pHeader := iq_stEntry.pRxBuffer;
IF pHeader = 0 THEN
	RETURN;
END_IF
IF pHeader^.DeviceCount=0 OR pHeader^.DeviceCount>iq_stEntry.nMaxRecords THEN RETURN; END_IF
IF pHeader^.DeviceCount>(nPayloadBytes-SIZEOF(ST_MqttCommandHeader))/iq_stEntry.nElementSize THEN RETURN; END_IF
nRequiredBytes:=SIZEOF(ST_MqttCommandHeader)+pHeader^.DeviceCount*iq_stEntry.nElementSize;
IF nRequiredBytes>nPayloadBytes THEN RETURN; END_IF
nRecords := pHeader^.DeviceCount;		// 버퍼에 들어갈 수만큼 (위 검사로 실제 받은 레코드 수 이하)
q_nReceived := nRecords;		// [STD 21번 수정 2026-11-09: 받은 레코드 수]

(* 1부터 셈: 레코드가 0개면 돌지 않음 (0 - 1을 UDINT로 계산하면 넘쳐서 약 42억 번 돌게 됨) *)
FOR k := 1 TO nRecords DO
	pRecord := iq_stEntry.pRxBuffer;
	pRecord := pRecord + SIZEOF(ST_MqttCommandHeader) + (k - 1) * iq_stEntry.nElementSize;

	IF iq_stEntry.bIndexed THEN
		pIndex := pRecord + iq_stEntry.nIndexOffset;	// DeviceIndex 위치 (command는 SequenceNumber 뒤 4 B, config는 맨 앞) [2026-11-12]
		IF pIndex^ >= DEVICE_ID_BASE + iq_stEntry.nDeviceIdBase THEN
			nDev := pIndex^ - DEVICE_ID_BASE - iq_stEntry.nDeviceIdBase;
		ELSE
			nDev := iq_stEntry.nDeviceCapacity;	// 범위 밖 → 버림
		END_IF
	ELSE
		nDev := 0;							// 단일 레코드 (protection)
	END_IF

	IF nDev < iq_stEntry.nDeviceCapacity THEN
		pDest := iq_stEntry.pDestArray;
		pDest := pDest + nDev * iq_stEntry.nElementSize;
		MEMCPY(destAddr := pDest, srcAddr := pRecord, n := iq_stEntry.nElementSize);
		F_MqttDistribute := F_MqttDistribute + 1;
	END_IF
END_FOR

END_FUNCTION

// ---- 20_Module/Mqtt/FB_MqttPublish.TcPOU
FUNCTION_BLOCK FB_MqttPublish		// MQTT 발행 (브로커 1개): 장치 토픽·config echo 토픽을 1 s마다 발행, 로거 이벤트는 M_PublishLogger로 1건씩
VAR_INPUT
	i_nSiteId		: UDINT;
	i_sConnLabel	: STRING(10);	// 연결 구분 ('Cloud', 'local', 'Azure'). ClientId에만 씀
	i_sHost			: STRING(15);
	i_nPort			: UINT;
	i_sUserName		: STRING;
	i_sUserPassword	: STRING;	// 접속 값은 첫 호출 때 한 번 읽음
	i_sInstance		: STRING(4) := '';	// ClientId 뒤에 붙임. 이중화: 두 PLC가 같은 ClientId로 접속하면 브로커가 서로 끊으므로 PLC마다 다르게 ('-P', '-S')
	i_bPublish		: BOOL := TRUE;	// FALSE = 접속은 유지하고 발행만 안 함 (이중화: Active만 발행)
	i_astDeviceTable	: ARRAY[1..GVL_MQTT.DEVICE_TOPIC_COUNT] OF ST_MqttPubEntry;	// 장치 토픽 표 (FB_MqttMain.A_InitPublishTable)
	i_astConfigTable	: ARRAY[1..GVL_MQTT.CONFIG_TOPIC_COUNT] OF ST_MqttPubEntry;	// config echo 토픽 표
END_VAR
VAR
	_sSiteId			: STRING;
	_sClientId			: STRING;
	_sHost				: STRING(15);
	_nPort				: UINT;
	_sUserName			: STRING;
	_sUserPassword		: STRING;
	_asDeviceTopic		: ARRAY[1..GVL_MQTT.DEVICE_TOPIC_COUNT] OF STRING(80);
	_asConfigTopic		: ARRAY[1..GVL_MQTT.CONFIG_TOPIC_COUNT] OF STRING(80);
	_sLoggerTopic		: STRING(80);
	_fbClient			: FB_IotMqttClient;
	_fbQueue			: FB_IotMqttMessageQueue;
	_i					: UINT;
	_bSetParameter		: BOOL := TRUE;
	_bConnect			: BOOL := TRUE;
	_bPublished			: BOOL;
	_tonPeriod			: TON := (PT := T#1S);		// 발행 주기
END_VAR

IF _bSetParameter THEN
	_bSetParameter := FALSE;
	_sSiteId		:= UDINT_TO_STRING(i_nSiteId);
	_sHost			:= i_sHost;
	_nPort			:= i_nPort;
	_sClientId		:= CONCAT(CONCAT('dgspms/pub-', i_sConnLabel), CONCAT('/', _sSiteId));
	_sClientId		:= CONCAT(_sClientId, i_sInstance);
	_sUserName		:= i_sUserName;
	_sUserPassword	:= i_sUserPassword;
	(* 장치 토픽: dgspms/{solution}/{site_id}/{device_name} *)
	FOR _i := 1 TO GVL_MQTT.DEVICE_TOPIC_COUNT DO
		_asDeviceTopic[_i] := CONCAT(CONCAT(CONCAT('dgspms/', GVL_MQTT.SOLUTION_NAME), CONCAT('/', _sSiteId)),
									CONCAT('/', i_astDeviceTable[_i].sTopic));
	END_FOR
	(* config echo 토픽: dgspms/{solution}/{site_id}/config/{device_name} *)
	FOR _i := 1 TO GVL_MQTT.CONFIG_TOPIC_COUNT DO
		_asConfigTopic[_i] := CONCAT(CONCAT(CONCAT('dgspms/', GVL_MQTT.SOLUTION_NAME), CONCAT('/', _sSiteId)),
									CONCAT(CONCAT('/', i_astConfigTable[_i].sCategory), CONCAT('/', i_astConfigTable[_i].sTopic)));
	END_FOR

	(* 로거 토픽: dgspms/{solution}/{site_id}/{LOGGER_TOPIC} (주기 발행 아님. M_PublishLogger로 이벤트가 생길 때만) *)
	_sLoggerTopic := CONCAT(CONCAT(CONCAT('dgspms/', GVL_MQTT.SOLUTION_NAME), CONCAT('/', _sSiteId)), CONCAT('/', GVL_MQTT.LOGGER_TOPIC));

	_fbClient.sClientId		:= _sClientId;
	_fbClient.sUserName		:= _sUserName;
	_fbClient.sUserPassword	:= _sUserPassword;
	_fbClient.sHostName		:= _sHost;
	_fbClient.nHostPort		:= _nPort;
	_fbClient.sTopicPrefix	:= '';
	_fbClient.ipMessageQueue := _fbQueue;
END_IF

_fbClient.Execute(_bConnect);

IF _fbClient.bConnected AND i_bPublish THEN
	_tonPeriod(IN := TRUE);
	IF _tonPeriod.Q THEN
		_tonPeriod(IN := FALSE);
		FOR _i := 1 TO GVL_MQTT.DEVICE_TOPIC_COUNT DO
			IF i_astDeviceTable[_i].nDeviceCount > 0 THEN
			_bPublished := _fbClient.Publish(sTopic := _asDeviceTopic[_i],
						pPayload := i_astDeviceTable[_i].pStaging,
						nPayloadSize := i_astDeviceTable[_i].nStagingSize,
						eQos := TcIotMqttQos.AtMostOnceDelivery,
						bRetain := FALSE,
						bQueue := FALSE);
			END_IF
		END_FOR
		FOR _i := 1 TO GVL_MQTT.CONFIG_TOPIC_COUNT DO
			IF i_astConfigTable[_i].nDeviceCount > 0 THEN
			_bPublished := _fbClient.Publish(sTopic := _asConfigTopic[_i],
						pPayload := i_astConfigTable[_i].pStaging,
						nPayloadSize := i_astConfigTable[_i].nStagingSize,
						eQos := TcIotMqttQos.AtMostOnceDelivery,
						bRetain := FALSE,
						bQueue := FALSE);
			END_IF
		END_FOR
	END_IF
END_IF

METHOD M_PublishLogger : BOOL		// 로거 이벤트 1건 발행 (QoS 1, 반복 없음). 접속돼 있고 보냈으면 TRUE (FB_MqttMain.A_PublishLogger가 부름)
VAR_INPUT
	i_pPayload	: PVOID;		// ST_LoggerPublish_V1
	i_nSize		: UDINT;
END_VAR
M_PublishLogger := FALSE;
IF _bSetParameter OR NOT _fbClient.bConnected OR NOT i_bPublish THEN
	RETURN;		// 아직 접속 전: 큐에 남아 있다가 접속하면 나감. 발행 허가 없음(이중화 대기)도 보내지 않음
END_IF
M_PublishLogger := _fbClient.Publish(sTopic := _sLoggerTopic,
						pPayload := i_pPayload,
						nPayloadSize := i_nSize,
						eQos := TcIotMqttQos.AtLeastOnceDelivery,
						bRetain := FALSE,
						bQueue := FALSE);
END_METHOD

END_FUNCTION_BLOCK

// ---- 20_Module/Mqtt/Logger/FB_MqttLoggerListener.TcPOU
FUNCTION_BLOCK FB_MqttLoggerListener EXTENDS FB_ListenerBase2		// 로거 리스너: TwinCAT 이벤트 로거에 남은 PMS 이벤트를 받아 시각·문구를 큐에 쌓음 (로거 토픽 발행용. FB_MqttMain이 M_Cycle·M_GetPacket을 부름)
(* - FB_EventLog가 이벤트 로거에 남긴 것을 그대로 받는다 (메시지 1회, 알람 발생·해소). 기록하는 곳은 FB_EventLog 하나이고, 이 FB는 받아서 옮기기만 한다
   - 받는 이벤트 클래스: PmsSystem·PmsProt·PmsOutput·PmsSeq (TwinCAT 시스템 이벤트는 받지 않음). 구독은 클래스 단위(TC_EVENT_CLASSES)
   - 제어기 TwinCAT 런타임 3.1.4024.17 이상 필요 (FB_ListenerBase2). 낮으면 구독이 16#98110701(서비스 미지원)로 실패해 아무것도 받지 못함 (_hrSubscribe)
   - 문구: FB_RequestEventText로 비동기로 받는다 (UTF-8 → F_Utf8ToWstring). 해소는 앞에 '[해소] '.
     LOGGER_TEXT_MAX(100)자를 넘으면 99자 + '…'로 자르고 q_nTruncated를 센다 (문구 규칙: 인자를 채운 로그 문구 95자 이내, PMS_STD.md 7장)
   - 시각: 로거 기록 시각(UTC)을 현지 시각으로 바꾼다 (i_nUtcOffset, FB_MqttMain이 계산). 시간대를 아직 모르면 기다린다
   - 큐: LOGGER_QUEUE칸 링 버퍼. 브로커마다 M_GetPacket으로 다음 번호를 꺼내 간다. 밀려서 덮어쓰인 것은 건너뛰고 q_nLost
   - 본체는 부르지 않는다 (리스너 기반 FB). 매 스캔 M_Cycle을 부른다 *)
VAR_OUTPUT
	q_bSubscribed	: BOOL;		// 이벤트 로거 구독 중
	q_nReceived		: UDINT;	// 받은 이벤트 수 (= 마지막 이벤트 번호)
	q_nTruncated	: UDINT;	// LOGGER_TEXT_MAX를 넘어 자른 수 (문구 규칙 위반: 문구 틀·인자를 줄일 것)
	q_nTextError	: UDINT;	// 문구를 못 받아 대체 문구를 쓴 수
	q_nLost			: UDINT;	// 브로커가 밀려 보내지 못하고 덮어쓰인 수 (브로커 합)
END_VAR
VAR CONSTANT
	TEXT_TIMEOUT	: ULINT := 50000000;	// 문구 요청 제한 5 s (100 ns 단위). 넘으면 대체 문구
	SUBSCRIBE_RETRY	: UINT := 100;			// 구독 실패 뒤 다시 시도까지 M_Cycle 호출 수 (MqttTask 10 ms × 100 = 1 s)
	CLEARED_MARK	: WSTRING(7) := "[해소] ";	// 알람 해소 표시 (5자)
END_VAR
VAR
	_fbFilter		: FB_TcEventFilter;
	_hrSubscribe	: HRESULT;
	_hrExecute		: HRESULT;
	_nSubscribeWait	: UINT;
	_nUtcOffset		: LINT;		// 현지 시각 − UTC (100 ns). M_Cycle 입력
	_bTimeValid		: BOOL;
	_nWriteNo		: UDINT;	// 마지막으로 넣은 이벤트 번호
	_astSlot		: ARRAY[1..GVL_MQTT.LOGGER_QUEUE] OF ST_LoggerSlot;
	_afbText		: ARRAY[1..GVL_MQTT.LOGGER_QUEUE] OF FB_RequestEventText;	// 칸마다 하나 (한 스캔에 여러 이벤트가 와도 요청이 겹치지 않게)
	{attribute 'TcEncoding' := 'UTF-8'}
	_sText			: STRING(511);		// 받은 문구 (UTF-8. 한글 95자 ≈ 285 byte)
	_wsText			: WSTRING(255);
	_k				: UINT;
	_nNow			: ULINT;
END_VAR

(* 본체는 쓰지 않는다. M_Cycle을 부른다 *)

METHOD M_Cycle		// 매 스캔 (MqttTask): 구독 → 이벤트 받기(콜백이 큐에 넣음) → 칸마다 문구·시각 채우기
VAR_INPUT
	i_nUtcOffset	: LINT;		// 현지 시각 − UTC (100 ns 단위)
	i_bTimeValid	: BOOL;		// i_nUtcOffset을 믿을 수 있음 (현지 시각을 얻음)
END_VAR
_nUtcOffset	:= i_nUtcOffset;
_bTimeValid	:= i_bTimeValid;

(* 1. 구독 (처음, 실패하면 SUBSCRIBE_RETRY 호출 뒤 다시) *)
IF NOT THIS^.bSubscribed THEN
	IF _nSubscribeWait = 0 THEN
		(* 클래스 단위 (TC_EVENT_CLASSES): 클래스 안의 이벤트를 추가·삭제·이름 변경해도 고치지 않음. 새 이벤트 클래스를 만들면 여기에 한 줄 *)
		_fbFilter.Clear().EventClass.EqualTo(TC_EVENT_CLASSES.PmsSystem)
			.OR_OP().EventClass.EqualTo(TC_EVENT_CLASSES.PmsProt)
			.OR_OP().EventClass.EqualTo(TC_EVENT_CLASSES.PmsOutput)
			.OR_OP().EventClass.EqualTo(TC_EVENT_CLASSES.PmsSeq);
		_hrSubscribe := THIS^.Subscribe2(_fbFilter);
		_nSubscribeWait := SUBSCRIBE_RETRY;
	ELSE
		_nSubscribeWait := _nSubscribeWait - 1;
	END_IF
END_IF
q_bSubscribed := THIS^.bSubscribed;

(* 2. 이벤트 받기: 이 안에서 OnMessageSent·OnAlarmRaised·OnAlarmCleared가 불려 큐에 넣고 문구를 요청함 *)
_hrExecute := THIS^.Execute();

(* 3. 칸마다: 문구가 오면 받고, 시간대를 알면 시각 문자열을 만들어 발행 준비 *)
_nNow := F_GetSystemTime();
FOR _k := 1 TO GVL_MQTT.LOGGER_QUEUE DO
	IF _astSlot[_k].bRequesting THEN
		IF _afbText[_k].bError OR (_nNow - _astSlot[_k].nRequestStart) > TEXT_TIMEOUT THEN
			q_nTextError := q_nTextError + 1;
			M_SetText(i_nSlot := _k, i_wsText := WCONCAT("로그 문구를 가져오지 못함: 이벤트 ID ", TO_WSTRING(_astSlot[_k].nEventId)));
		ELSIF NOT _afbText[_k].bBusy THEN
			_sText := '';
			_afbText[_k].GetString(_sText, SIZEOF(_sText));
			M_SetText(i_nSlot := _k, i_wsText := F_Utf8ToWstring(i_pSrc := ADR(_sText), i_nSrcSize := SIZEOF(_sText)));
		END_IF
	END_IF
	IF _astSlot[_k].bTextDone AND NOT _astSlot[_k].bReady AND _bTimeValid THEN
		_astSlot[_k].sTime	:= M_TimeText(_astSlot[_k].nTimestamp);
		_astSlot[_k].bReady	:= TRUE;
	END_IF
END_FOR
END_METHOD

METHOD M_GetPacket : BOOL		// 브로커 하나가 보낼 다음 이벤트 패킷. TRUE면 iq_stPacket을 채움 (보낸 뒤 부르는 쪽이 iq_nNext를 1 올림)
VAR_INPUT
	i_nSiteId	: UDINT;
END_VAR
VAR_IN_OUT
	iq_nNext	: UDINT;				// 이 브로커가 다음에 보낼 이벤트 번호 (1부터)
	iq_stPacket	: ST_LoggerPublish_V1;
END_VAR
VAR
	k			: UINT;
	nOldest		: UDINT;
	nBytes		: UDINT;
END_VAR
M_GetPacket := FALSE;
IF iq_nNext = 0 THEN
	iq_nNext := 1;
END_IF
IF _nWriteNo < iq_nNext THEN
	RETURN;		// 새 이벤트 없음
END_IF

(* 큐 칸 수보다 많이 밀렸으면 덮어쓰인 것은 건너뜀 *)
IF _nWriteNo - iq_nNext >= UINT_TO_UDINT(GVL_MQTT.LOGGER_QUEUE) THEN
	nOldest		:= _nWriteNo - UINT_TO_UDINT(GVL_MQTT.LOGGER_QUEUE) + 1;
	q_nLost		:= q_nLost + (nOldest - iq_nNext);
	iq_nNext	:= nOldest;
END_IF

k := M_SlotOf(iq_nNext);
IF _astSlot[k].nNo <> iq_nNext OR NOT _astSlot[k].bReady THEN
	RETURN;		// 문구·시각을 아직 받는 중
END_IF

(* 매번 비우고 채움: 짧은 문구의 null 뒤에 지난 문구가 남지 않게.
   문자열은 대입(:=)하지 않고 길이 + null만 MEMCPY: 문자열 대입은 선언 크기 전체를 복사해서,
   큐 칸을 돌려 쓰는 동안 null 뒤에 남은 옛 문구까지 패킷에 들어감 (PC 도구 재pack 비교에서 "불일치"로 보임) *)
MEMSET(destAddr := ADR(iq_stPacket), fillByte := 0, n := SIZEOF(iq_stPacket));
iq_stPacket.Header.HeaderVersion	:= GVL_MQTT.HEADER_VERSION;
iq_stPacket.Header.DeviceVersion	:= GVL_MQTT.LOGGER_VERSION;
iq_stPacket.Header.SiteId			:= i_nSiteId;
nBytes := INT_TO_UDINT(LEN(_astSlot[k].sTime)) + 1;
IF nBytes > SIZEOF(iq_stPacket.Header.TimeStamp) THEN
	nBytes := SIZEOF(iq_stPacket.Header.TimeStamp);
END_IF
MEMCPY(destAddr := ADR(iq_stPacket.Header.TimeStamp), srcAddr := ADR(_astSlot[k].sTime), n := nBytes);
nBytes := (INT_TO_UDINT(WLEN(_astSlot[k].wsText)) + 1) * 2;
IF nBytes > SIZEOF(iq_stPacket.Contents) THEN
	nBytes := SIZEOF(iq_stPacket.Contents);
END_IF
MEMCPY(destAddr := ADR(iq_stPacket.Contents), srcAddr := ADR(_astSlot[k].wsText), n := nBytes);
M_GetPacket := TRUE;
END_METHOD

METHOD OnMessageSent : HRESULT		// 메시지 1건 (FB_LogMsg) → 큐
VAR_INPUT
	fbEvent	: REFERENCE TO FB_TcEvent;
END_VAR
M_Push(i_fbEvent := fbEvent, i_bCleared := FALSE);
OnMessageSent := S_OK;		// S_OK여야 이번 스캔에 다음 콜백을 계속 받음
END_METHOD

METHOD OnAlarmRaised : HRESULT		// 알람 발생 (FB_LogAlarm) → 큐
VAR_INPUT
	fbEvent	: REFERENCE TO FB_TcEvent;
END_VAR
M_Push(i_fbEvent := fbEvent, i_bCleared := FALSE);
OnAlarmRaised := S_OK;		// S_OK여야 이번 스캔에 다음 콜백을 계속 받음
END_METHOD

METHOD OnAlarmCleared : HRESULT		// 알람 해소 → 큐 ('[해소] ' 표시)
VAR_INPUT
	fbEvent	: REFERENCE TO FB_TcEvent;
END_VAR
M_Push(i_fbEvent := fbEvent, i_bCleared := TRUE);
OnAlarmCleared := S_OK;		// S_OK여야 이번 스캔에 다음 콜백을 계속 받음
END_METHOD

METHOD OnAlarmConfirmed : HRESULT		// 쓰지 않음
VAR_INPUT
	fbEvent	: REFERENCE TO FB_TcEvent;
END_VAR
OnAlarmConfirmed := S_OK;		// 확인(Confirm)은 쓰지 않음 (알람을 확인 없이 만듦)
END_METHOD

METHOD PRIVATE M_Push		// 받은 이벤트를 큐 다음 칸에 넣고 문구를 요청 (콜백이 부름). 큐가 차면 가장 오래된 칸을 덮어씀
VAR_INPUT
	i_fbEvent	: REFERENCE TO FB_TcEvent;
	i_bCleared	: BOOL;
END_VAR
VAR
	k			: UINT;
END_VAR
_nWriteNo	:= _nWriteNo + 1;
q_nReceived	:= _nWriteNo;
k := M_SlotOf(_nWriteNo);

_astSlot[k].nNo				:= _nWriteNo;
_astSlot[k].nTimestamp		:= i_fbEvent.nTimestamp;
_astSlot[k].nEventId		:= i_fbEvent.nEventId;
_astSlot[k].bCleared		:= i_bCleared;
_astSlot[k].bRequesting		:= TRUE;
_astSlot[k].nRequestStart	:= F_GetSystemTime();
_astSlot[k].bTextDone		:= FALSE;
_astSlot[k].bReady			:= FALSE;
_astSlot[k].sTime			:= '';
_astSlot[k].wsText			:= "";

(* 문구는 비동기로 옴 (M_Cycle에서 받음). 인자는 요청할 때 넘김 (콜백 밖에서는 i_fbEvent를 쓸 수 없음) *)
_afbText[k].Request(eventClass := i_fbEvent.EventClass, nEventId := i_fbEvent.nEventId,
					nLangId := GVL_MQTT.LOGGER_LANG_ID, ipArgs := i_fbEvent.ipArguments);
END_METHOD

METHOD PRIVATE M_SetText		// 받은 문구를 칸에 넣음: 해소 표시를 붙이고 LOGGER_TEXT_MAX자로 맞춤
VAR_INPUT
	i_nSlot		: UINT;
	i_wsText	: WSTRING(255);
END_VAR
_wsText := i_wsText;
IF _astSlot[i_nSlot].bCleared THEN
	_wsText := WCONCAT(CLEARED_MARK, _wsText);
END_IF
IF WLEN(_wsText) > GVL_MQTT.LOGGER_TEXT_MAX THEN
	_wsText := WCONCAT(WLEFT(_wsText, GVL_MQTT.LOGGER_TEXT_MAX - 1), "…");
	q_nTruncated := q_nTruncated + 1;
END_IF
_astSlot[i_nSlot].wsText		:= _wsText;
_astSlot[i_nSlot].bRequesting	:= FALSE;
_astSlot[i_nSlot].bTextDone		:= TRUE;
END_METHOD

METHOD PRIVATE M_SlotOf : UINT		// 이벤트 번호 → 큐 칸 (1..LOGGER_QUEUE)
VAR_INPUT
	i_nNo	: UDINT;
END_VAR
M_SlotOf := UDINT_TO_UINT(((i_nNo - 1) MOD UINT_TO_UDINT(GVL_MQTT.LOGGER_QUEUE)) + 1);
END_METHOD

METHOD PRIVATE M_TimeText : STRING(23)		// 로거 시각(FILETIME, UTC) → 현지 시각 문자열
VAR_INPUT
	i_nFileTime	: ULINT;
END_VAR
VAR
	nLocal		: ULINT;
	stFileTime	: T_FILETIME;
END_VAR
nLocal := LINT_TO_ULINT(ULINT_TO_LINT(i_nFileTime) + _nUtcOffset);
MEMCPY(destAddr := ADR(stFileTime), srcAddr := ADR(nLocal), n := SIZEOF(stFileTime));
M_TimeText := F_MqttTimeText(FILETIME_TO_SYSTEMTIME(stFileTime));
END_METHOD

END_FUNCTION_BLOCK

// ---- 20_Module/Mqtt/Logger/F_Utf8ToWstring.TcPOU
FUNCTION F_Utf8ToWstring : WSTRING(255)		// UTF-8 바이트(0에서 끝남) → WSTRING(UTF-16). 255자에서 자름. 4바이트 문자(이모지 등)·잘못된 바이트는 U+FFFD 한 글자
(* 이벤트 로거 문구(FB_RequestEventText.GetString)는 UTF-8 STRING으로만 받을 수 있어서 쓴다.
   한글(U+AC00~)은 UTF-8 3바이트 → UTF-16 한 칸 *)
VAR_INPUT
	i_pSrc		: PVOID;				// UTF-8 문자열 시작 주소 (STRING 변수의 ADR)
	i_nSrcSize	: UDINT;				// 그 버퍼 크기 (byte, SIZEOF). 0을 만나면 그 앞에서 끝
END_VAR
VAR CONSTANT
	MAX_SRC		: UDINT := 1024;		// 읽는 최대 바이트
	MAX_CHARS	: UINT := 255;
	BAD_CHAR	: WORD := 16#FFFD;
END_VAR
VAR
	pSrc		: POINTER TO ARRAY[0..1023] OF BYTE;	// MAX_SRC
	wsOut		: WSTRING(255);
	pOut		: POINTER TO ARRAY[0..255] OF WORD;		// wsOut (MAX_CHARS + null)
	nSize		: UDINT;
	i			: UDINT;
	nChars		: UINT;
	nLen		: UDINT;
	b0			: BYTE;
	b1			: BYTE;
	b2			: BYTE;
	wChar		: WORD;
END_VAR

F_Utf8ToWstring := "";
IF i_pSrc = 0 THEN
	RETURN;
END_IF
pSrc	:= i_pSrc;
pOut	:= ADR(wsOut);
nSize	:= MIN(i_nSrcSize, MAX_SRC);
i		:= 0;
nChars	:= 0;

WHILE i < nSize AND nChars < MAX_CHARS DO
	b0 := pSrc^[i];
	IF b0 = 0 THEN
		EXIT;
	END_IF
	wChar	:= BAD_CHAR;
	nLen	:= 1;
	IF b0 < 16#80 THEN							// 1바이트 (ASCII)
		wChar := BYTE_TO_WORD(b0);
	ELSIF (b0 AND 16#E0) = 16#C0 THEN			// 2바이트
		IF i + 1 < nSize THEN
			b1 := pSrc^[i + 1];
			IF (b1 AND 16#C0) = 16#80 THEN
				wChar	:= SHL(BYTE_TO_WORD(b0 AND 16#1F), 6) OR BYTE_TO_WORD(b1 AND 16#3F);
				nLen	:= 2;
			END_IF
		END_IF
	ELSIF (b0 AND 16#F0) = 16#E0 THEN			// 3바이트 (한글 등)
		IF i + 2 < nSize THEN
			b1 := pSrc^[i + 1];
			b2 := pSrc^[i + 2];
			IF (b1 AND 16#C0) = 16#80 AND (b2 AND 16#C0) = 16#80 THEN
				wChar	:= SHL(BYTE_TO_WORD(b0 AND 16#0F), 12) OR SHL(BYTE_TO_WORD(b1 AND 16#3F), 6) OR BYTE_TO_WORD(b2 AND 16#3F);
				nLen	:= 3;
			END_IF
		END_IF
	ELSIF (b0 AND 16#F8) = 16#F0 THEN			// 4바이트 → U+FFFD 한 글자
		nLen := 4;
	END_IF
	pOut^[nChars]	:= wChar;
	nChars			:= nChars + 1;
	i				:= i + nLen;
END_WHILE
pOut^[nChars] := 0;
F_Utf8ToWstring := wsOut;

END_FUNCTION

// ---- 20_Module/Mqtt/F_MqttTimeText.TcPOU
FUNCTION F_MqttTimeText : STRING(23)		// 시각 → 'YYYY-MM-DD hh:mm:ss.xxx' (MQTT 헤더 TimeStamp 형식, 23자). FB_MqttMain(발행 헤더)·FB_MqttLoggerListener(로거 시각)가 같이 씀
VAR_INPUT
	i_stTime	: TIMESTRUCT;
END_VAR

(* Tc2_Utilities SYSTEMTIME_TO_STRING 형식은 'YYYY-MM-DD-hh:mm:ss.xxx' → 11번째 글자 '-'를 공백으로 *)
F_MqttTimeText := REPLACE(SYSTEMTIME_TO_STRING(i_stTime), ' ', 1, 11);

END_FUNCTION

// ---- 20_Module/Mqtt/FB_EmsCommand.TcPOU
FUNCTION_BLOCK FB_EmsCommand		// 명령 핸들러 (MqttTask): 받은 EMS command 레코드 → Std 명령 (PCS·BMS 상태 명령, 충전·방전 P 지령)
(* - 받은 레코드의 CommandType이 0이 아니면 한 번 해석하고 0으로 지운다 (같은 레코드를 다시 실행하지 않음)
   - 새 명령마다 번호(nSeq, anPcsPSeq)를 1 올린다. 받는 쪽(FB_SrcEms)은 번호 변화로 새 명령을 안다
   - 결과 q_stCmd는 지금까지 받은 명령 전체(마지막 값 유지). 바뀐 스캔에만 q_bChanged가 켜지고, PRG_Mqtt가 GVL_IF에 올린다
   - 받은 레코드 배열은 0부터 (GVL_MQTT 수신 배열 칸 = 레코드 DeviceIndex − 1, F_MqttDistribute.DEVICE_ID_BASE = 1). 결과는 Std 규칙대로 1부터 (칸 = DeviceIndex)
   - 이상한 값(NaN·무한대·절댓값이 MAX_VALUE 초과)의 P 지령은 버리고 센다. NaN은 비교하면 PLC가 멈추므로 F_IsFinite(비트)로 먼저 거른다. 정격 대비 상한은 코어 명령 필터(g_stCmdFilter)가 다시 거른다
   PCS CommandType: 1 Run, 2 Stop, 3 Standby, 4 충전(Value kW), 5 방전(Value kW), 6 비상정지, 7 리셋
   BAT CommandType: 1 접촉기 투입(Close), 2 개방(Open), 3 비상정지, 4 리셋, 11 랙 컨택터 닫기, 12 랙 컨택터 열기 (Value = 랙 번호 1~)
   5 시스템(랙 전체 40013) 연결, 6 차단, 7 충전 컨택터(40014) 닫기, 8 열기, 9 방전 컨택터(40015) 닫기, 10 열기 → astBatCtl [2026-11-13]
   (인터페이스 100.Command) *)
VAR_INPUT
	i_nRxCount			: UDINT;	// command 메시지 수신 누계 (브로커 3개 합)
END_VAR
VAR_IN_OUT
	iq_astPcsCommand	: ARRAY[0..GVL_PARAM.PCS_COUNT-1] OF ST_MqttCommand_Rx;	// GVL_MQTT.g_astPcsCommand
	iq_astBatCommand	: ARRAY[0..GVL_PARAM.BMS_COUNT-1] OF ST_MqttCommand_Rx;	// GVL_MQTT.g_astBatCommand
END_VAR
VAR_OUTPUT
	q_stCmd				: ST_IfEmsCmd;	// 지금까지 받은 명령
	q_bChanged			: BOOL;			// 이번 스캔에 q_stCmd가 바뀜
	q_nUnknownCount		: UDINT;		// 모르는 CommandType을 받은 횟수
	q_nBadValueCount	: UDINT;		// 이상한 값의 P 지령을 버린 횟수
END_VAR
VAR CONSTANT
	MAX_VALUE			: REAL := 1.0E7;	// kW. 이보다 크면 이상값
END_VAR
VAR
	_i					: UINT;
	_n					: UINT;
	_ePcsCmd			: E_PcsCmd;
	_eBatCmd			: E_BatCmd;
	_bP					: BOOL;
	_fP					: REAL;
	_bValueOk			: BOOL;		// 받은 Value가 보통 숫자 (NaN·무한대 아님)
END_VAR

q_bChanged := FALSE;

// 명령이 없는 메시지도 '살아 있음'으로 셈
IF i_nRxCount <> q_stCmd.nRxCount THEN
	q_stCmd.nRxCount := i_nRxCount;
	q_bChanged := TRUE;
END_IF

(* PCS *)
FOR _i := 0 TO GVL_PARAM.PCS_COUNT - 1 DO
	IF iq_astPcsCommand[_i].CommandType <> 0 THEN
		_n := _i + 1;
		_ePcsCmd	:= E_PcsCmd.None;
		_bP			:= FALSE;
		_bValueOk	:= F_IsFinite(iq_astPcsCommand[_i].Value);	// NaN은 크기 비교·ABS 전에 비트로 거름 (비교하면 PLC가 멈춤)
		CASE iq_astPcsCommand[_i].CommandType OF
			1:	_ePcsCmd := E_PcsCmd.Run;
			2:	_ePcsCmd := E_PcsCmd.Stop;
			3:	_ePcsCmd := E_PcsCmd.Standby;
			4:	_bP := TRUE;	IF _bValueOk THEN _fP := -ABS(iq_astPcsCommand[_i].Value); END_IF	// 충전
			5:	_bP := TRUE;	IF _bValueOk THEN _fP := ABS(iq_astPcsCommand[_i].Value); END_IF		// 방전
			6:	_ePcsCmd := E_PcsCmd.EStop;
			7:	_ePcsCmd := E_PcsCmd.Reset;
		ELSE
			q_nUnknownCount := q_nUnknownCount + 1;
		END_CASE
		// P 지령 값 거르기: 보통 숫자가 아니거나 너무 크면 버림 (크기 비교는 보통 숫자일 때만)
		IF _bP THEN
			IF NOT _bValueOk THEN
				_bP := FALSE;
				q_nBadValueCount := q_nBadValueCount + 1;
			ELSIF ABS(iq_astPcsCommand[_i].Value) > MAX_VALUE THEN
				_bP := FALSE;
				q_nBadValueCount := q_nBadValueCount + 1;
			END_IF
		END_IF
		IF _ePcsCmd <> E_PcsCmd.None THEN
			q_stCmd.astPcs[_n].eCmd := _ePcsCmd;
			q_stCmd.astPcs[_n].nSeq := q_stCmd.astPcs[_n].nSeq + 1;
			q_bChanged := TRUE;
		END_IF
		IF _bP THEN
			q_stCmd.afPcsP[_n]		:= _fP;
			q_stCmd.anPcsPSeq[_n]	:= q_stCmd.anPcsPSeq[_n] + 1;
			q_bChanged := TRUE;
		END_IF
		iq_astPcsCommand[_i].CommandType := 0;		// 처리 완료
	END_IF
END_FOR

(* BAT (BMS) *)
FOR _i := 0 TO GVL_PARAM.BMS_COUNT - 1 DO
	IF iq_astBatCommand[_i].CommandType <> 0 THEN
		_n := _i + 1;
		_eBatCmd := E_BatCmd.None;
		CASE iq_astBatCommand[_i].CommandType OF
			1:	_eBatCmd := E_BatCmd.Close;
			2:	_eBatCmd := E_BatCmd.Open;
			3:	_eBatCmd := E_BatCmd.EStop;
			4:	_eBatCmd := E_BatCmd.Reset;
			5..10:	// 컨택터 하나씩 (FB_BmsContactorCommand가 번호를 해석) [2026-11-13]
				q_stCmd.astBatCtl[_n].nSeq := q_stCmd.astBatCtl[_n].nSeq + 1;
				q_stCmd.astBatCtl[_n].nType := UDINT_TO_UINT(iq_astBatCommand[_i].CommandType);
				q_bChanged := TRUE;
			11, 12:	// 랙 컨택터 닫기·열기. Value = 랙 번호 (정수가 아니거나 범위 밖이면 0 → FB_BmsRackCommand가 거절)
				q_stCmd.astBatRack[_n].nSeq := q_stCmd.astBatRack[_n].nSeq + 1;
				q_stCmd.astBatRack[_n].bClose := iq_astBatCommand[_i].CommandType = 11;
				IF iq_astBatCommand[_i].Value >= 1.0 AND iq_astBatCommand[_i].Value <= 16.0
					AND iq_astBatCommand[_i].Value = UINT_TO_REAL(REAL_TO_UINT(iq_astBatCommand[_i].Value)) THEN
					q_stCmd.astBatRack[_n].nRack := REAL_TO_UINT(iq_astBatCommand[_i].Value);
				ELSE
					q_stCmd.astBatRack[_n].nRack := 0;
				END_IF
				q_bChanged := TRUE;
		ELSE
			q_nUnknownCount := q_nUnknownCount + 1;
		END_CASE
		IF _eBatCmd <> E_BatCmd.None THEN
			q_stCmd.astBat[_n].eCmd := _eBatCmd;
			q_stCmd.astBat[_n].nSeq := q_stCmd.astBat[_n].nSeq + 1;
			q_bChanged := TRUE;
		END_IF
		iq_astBatCommand[_i].CommandType := 0;		// 처리 완료
	END_IF
END_FOR

END_FUNCTION_BLOCK

// ---- 10_Core/02_Util/F_IsFinite.TcPOU
FUNCTION F_IsFinite : BOOL		// 실수가 보통 숫자인가 (NaN·무한대가 아님). 비트로만 봄
// NaN을 크기 비교(<, >, <=, >=)하면 부동소수점 예외(SSE invalid operation)로 PLC가 멈춤 → 바깥에서 온 실수는 비교하기 전에 이것으로 먼저 거름
VAR_INPUT
	i_fValue	: REAL;
END_VAR
VAR
	pBits		: POINTER TO DWORD;
END_VAR

pBits := ADR(i_fValue);
F_IsFinite := (pBits^ AND 16#7F800000) <> 16#7F800000;		// 지수 비트가 모두 1이면 NaN 또는 무한대

END_FUNCTION

// ---- 20_Module/Mqtt/FB_EmsCmdGate.TcPOU
FUNCTION_BLOCK FB_EmsCmdGate		// EMS command 레코드 앞단: 같은 SequenceNumber 버리기 + Delay(ms)만큼 기다렸다가 내보내기
(* EMS command 레코드 중복 방지·지연 실행 (⑤출력 앞단 / 장치: PCS·BAT·UPS 명령 공통). 2026-11-12.
   기반 없음(신규).
   변경: 없음
   부호·단위: Delay ms. 명세: C:\gil\UPS\명세서\UPS_명세서.md WR-CMD-01, 인터페이스 100.Command (SequenceNumber·Delay)
   - 수신 배열(GVL_MQTT.g_ast*Command, 칸 = DeviceIndex-1)을 그대로 받아, 명령 핸들러(FB_EmsCommand, PRG_Mqtt UPS 칸)보다 먼저 부른다
   - 새 레코드(CommandType<>0)의 SequenceNumber가 그 칸에서 마지막으로 받은 번호와 같으면 버린다 (0은 거르지 않음)
   - Delay = 0이면 그대로 두어 이번 스캔에 처리된다. Delay > 0이면 레코드를 빼서 보관하고, 시간이 되면 그 칸에 다시 넣는다
   - 보관 중에 같은 칸에 새 명령이 오면 보관한 명령은 버리고 새 명령을 따른다 (마지막 명령이 우선)
   - Delay가 MAX_DELAY_MS를 넘으면 버린다
   - 재시작하면 마지막 번호와 보관 명령은 없어진다 (보관 중이던 명령은 실행하지 않음) *)
VAR_IN_OUT
	iq_astRec			: ARRAY[*] OF ST_MqttCommand_Rx;	// 수신 배열 (0부터, 칸 = DeviceIndex-1)
END_VAR
VAR_OUTPUT
	q_nDupCount			: UDINT;	// 같은 SequenceNumber라 버린 수
	q_nDelayedCount		: UDINT;	// Delay 때문에 보관한 수
	q_nReplacedCount	: UDINT;	// 보관 중 새 명령이 와서 버린 보관 명령 수
	q_nBadDelayCount	: UDINT;	// Delay가 너무 커서 버린 수
	q_nPendingCount		: UDINT;	// 지금 보관 중인 명령 수
END_VAR
VAR CONSTANT
	MAX_SLOTS			: DINT := 16;			// 다룰 수 있는 칸 수 (PCS·BMS·UPS 대수보다 커야 함)
	MAX_DELAY_MS		: UDINT := 3600000;		// 1시간
END_VAR
VAR
	_anLastSeq			: ARRAY[0..15] OF UDINT;
	_astPend			: ARRAY[0..15] OF ST_MqttCommand_Rx;
	_abPend				: ARRAY[0..15] OF BOOL;
	_atStart			: ARRAY[0..15] OF TIME;
	_tNow				: TIME;
	_i					: DINT;
	_s					: DINT;
END_VAR

_tNow := TIME();
q_nPendingCount := 0;
FOR _i := LOWER_BOUND(iq_astRec, 1) TO UPPER_BOUND(iq_astRec, 1) DO
	_s := _i - LOWER_BOUND(iq_astRec, 1);
	IF _s >= MAX_SLOTS THEN
		EXIT;
	END_IF
	IF iq_astRec[_i].CommandType <> 0 THEN
		IF iq_astRec[_i].SequenceNumber <> 0 AND iq_astRec[_i].SequenceNumber = _anLastSeq[_s] THEN
			iq_astRec[_i].CommandType := 0;		// 같은 명령이 다시 옴
			q_nDupCount := q_nDupCount + 1;
		ELSE
			_anLastSeq[_s] := iq_astRec[_i].SequenceNumber;
			IF _abPend[_s] THEN
				_abPend[_s] := FALSE;			// 새 명령이 기다리던 명령을 대신함
				q_nReplacedCount := q_nReplacedCount + 1;
			END_IF
			IF iq_astRec[_i].Delay > MAX_DELAY_MS THEN
				iq_astRec[_i].CommandType := 0;
				q_nBadDelayCount := q_nBadDelayCount + 1;
			ELSIF iq_astRec[_i].Delay > 0 THEN
				_astPend[_s] := iq_astRec[_i];
				_abPend[_s] := TRUE;
				_atStart[_s] := _tNow;
				iq_astRec[_i].CommandType := 0;	// 시간이 될 때까지 핸들러가 못 보게 함
				q_nDelayedCount := q_nDelayedCount + 1;
			END_IF
		END_IF
	ELSIF _abPend[_s] AND (_tNow - _atStart[_s]) >= UDINT_TO_TIME(_astPend[_s].Delay) THEN
		iq_astRec[_i] := _astPend[_s];			// 시간이 됨: 이번 스캔에 핸들러가 처리
		iq_astRec[_i].Delay := 0;
		_abPend[_s] := FALSE;
	END_IF
	IF _abPend[_s] THEN
		q_nPendingCount := q_nPendingCount + 1;
	END_IF
END_FOR

END_FUNCTION_BLOCK

// ---- 20_Module/Mqtt/PRG_PublishDeviceNo.TcPOU
PROGRAM PRG_PublishDeviceNo		// 발행 패킷 장치 번호·랙 소속·모듈 수 채우기: 모든 장치 번호(DeviceIndex·BatIndex·RackIndex·DeviceId) = 1부터 순번. 배열 칸은 0부터(메시지 안의 몇 번째 레코드) [1부터 2026-11-10] (PRG_Mqtt가 부름)
(* DB 키: PcsLog·BatLog는 DeviceIndex, RackLog는 DeviceIndex로 UNIQUE(TimeStamp, 장치키) 저장·조회한다.
   번호가 비면(모두 0) 1분 회차의 두 번째 장치부터 INSERT가 실패하므로 측정값과 따로 항상 채운다.
   측정값은 보고 매핑(FB_Report, 인터페이스 확정 후)이 채운다 *)
VAR
	i		: UINT;
END_VAR

FOR i := 0 TO GVL_PARAM.PCS_COUNT - 1 DO
	g_stPcsPublish.Devices[i].DeviceIndex := UINT_TO_UDINT(i + 1);
END_FOR

FOR i := 0 TO GVL_PARAM.BMS_COUNT - 1 DO
	g_stBatPublish.Devices[i].DeviceIndex := UINT_TO_UDINT(i + 1);
	g_astBatConfig[i].DeviceId := UINT_TO_UDINT(i + 1);
END_FOR

FOR i := 0 TO GVL_PARAM.RACK_COUNT - 1 DO
	g_stRackPublish.Devices[i].DeviceIndex := UINT_TO_UDINT(i + 1);
	// 소속·수량은 측정값이 아닌 시험 구성 메타데이터. 더미 발행을 꺼도 번호와 함께 유지한다.
	g_stRackPublish.Devices[i].BatIndex := UINT_TO_UDINT(i / GVL_PARAM.RACKS_PER_BMS + 1);
	g_stRackPublish.Devices[i].ModuleCount := UINT_TO_UDINT(GVL_PARAM.MODULES_PER_RACK);
END_FOR
FOR i:=0 TO GVL_PARAM.UPS_COUNT-1 DO
 g_stUpsPublish.Devices[i].DeviceIndex:=UINT_TO_UDINT(i+1); // UPS는 1부터
 g_astUpsConfig[i].DeviceId:=UINT_TO_UDINT(i+1);
 // Scaffold is not a measurement mapping: mark unavailable, and keep publish gate FALSE.
 g_stUpsPublish.Devices[i].Status:=1;
END_FOR
FOR i:=0 TO GVL_PARAM.BMS_COUNT-1 DO
 g_stBatPublish.Devices[i].Status:=1;
END_FOR
FOR i:=0 TO GVL_PARAM.RACK_COUNT-1 DO
 g_stRackPublish.Devices[i].Status:=1;
END_FOR
FOR i:=0 TO GVL_PARAM.BAT_MODULE_COUNT-1 DO
 g_stModulePublish.Devices[i].BatIndex:=UINT_TO_UDINT(i / (GVL_PARAM.RACKS_PER_BMS * GVL_PARAM.MODULES_PER_RACK) + 1);
 g_stModulePublish.Devices[i].RackIndex:=UINT_TO_UDINT((i / GVL_PARAM.MODULES_PER_RACK) MOD GVL_PARAM.RACKS_PER_BMS + 1);
 g_stModulePublish.Devices[i].DeviceIndex:=UINT_TO_UDINT(i MOD GVL_PARAM.MODULES_PER_RACK + 1);
END_FOR
// 값을 채우는 매핑이 없는 토픽도 번호는 1부터 [1부터 2026-11-10]
g_stPmsPublish.Devices[0].DeviceIndex := 1;
FOR i:=0 TO GVL_PARAM.PV_COUNT-1 DO g_stPvPublish.Devices[i].DeviceIndex:=UINT_TO_UDINT(i + 1); END_FOR
FOR i:=0 TO GVL_PARAM.ESS_COUNT-1 DO g_stEssPublish.Devices[i].DeviceIndex:=UINT_TO_UDINT(i + 1); END_FOR
FOR i:=0 TO GVL_PARAM.TEMP_COUNT-1 DO g_stTempPublish.Devices[i].DeviceIndex:=UINT_TO_UDINT(i + 1); END_FOR
FOR i:=0 TO GVL_PARAM.AIR_CONDITIONER_COUNT-1 DO g_stAirConditionerPublish.Devices[i].DeviceIndex:=UINT_TO_UDINT(i + 1); END_FOR
FOR i:=0 TO GVL_PARAM.IMD_COUNT-1 DO g_stImdPublish.Devices[i].DeviceIndex:=UINT_TO_UDINT(i + 1); g_stImdPublish.Devices[i].Status:=1; END_FOR // 매핑이 채우기 전에는 통신 이상
FOR i:=0 TO GVL_PARAM.FIRE_COUNT-1 DO g_stFirePublish.Devices[i].DeviceIndex:=UINT_TO_UDINT(i + 1); g_stFirePublish.Devices[i].Status:=1; END_FOR // 매핑이 채우기 전에는 통신 이상

END_PROGRAM

// ---- 20_Module/Virtual/PRG_MqttTestData.TcPOU
PROGRAM PRG_MqttTestData		// 시험 전용 더미 발행 값 + 수신 기록 (PRG_Mqtt가 GVL_SITE.TEST_MODE일 때만 부름. 현장 빌드는 Virtual 폴더와 함께 뺌)
VAR
	bEnable			: BOOL := TRUE;			// FALSE면 더미 값을 쓰지 않음 (마지막 값 유지)
	tonUpdate		: TON := (PT := T#1S);	// 갱신 주기
	bFirstDone		: BOOL;					// 시작 직후 한 번은 바로 채움
	nTick			: UDINT;				// 갱신 횟수 (1 s마다 +1)
	fWave			: REAL;					// 삼각파 -1 ~ +1 (WAVE_PERIOD 초 주기)
	nHeartbeat		: UDINT;				// 0 ~ 99 반복 (BAT Heartbeat)
	fPcsP			: REAL;					// PCS 1대 유효전력 kW (방전 +)
	fBatSoc			: REAL;					// BAT SOC %
	fDev			: REAL;					// 장치 번호 (실수)
	nRacksPerBat	: UINT;					// BAT 1대에 속한 랙 수
	afPvEnergy		: ARRAY[0..GVL_PARAM.PV_COUNT-1] OF REAL;		// PV 누적 발전량 kWh
	afEssEnergy		: ARRAY[0..GVL_PARAM.ESS_COUNT-1] OF REAL;		// ESS 누적 방전량 kWh
	afEssEnergyRev	: ARRAY[0..GVL_PARAM.ESS_COUNT-1] OF REAL;		// ESS 누적 충전량 kWh
	fP				: REAL;
	i				: UINT;

	(* ---------- 수신 시험 핸들러 A_HandleRx (PRG_Mqtt가 FB_MqttMain 다음, 명령 핸들러 FB_EmsCommand 앞에서 부름) ----------
	   - 새 수신 판별은 v3_1과 같은 타임스탬프 방식: FB_MqttSubscribe가 헤더 TimeStamp가 바뀐 메시지만 q_an???RxCount +1
	     → EMS는 메시지마다 헤더 TimeStamp를 바꿔 보내야 새 수신으로 셈
	   - 브로커별 2중 배열 [1 Cloud, 2 Local, 3 Azure, 토픽]. command 토픽 1 pcs, 2 bat / config 토픽 1 pcs, 2 bat, 3 protection
	   - 받은 레코드는 FB_EmsCommand가 CommandType을 0으로 지우기 전에 사본으로 남김 *)
	anBrokerCmdCount	: ARRAY[1..3, 1..GVL_MQTT.COMMAND_TOPIC_COUNT] OF UDINT;		// 브로커별 command 수신 횟수 (FB_MqttSubscribe.q_anCmdRxCount)
	asBrokerCmdTime		: ARRAY[1..3, 1..GVL_MQTT.COMMAND_TOPIC_COUNT] OF STRING(23);	// 브로커별 마지막 command 헤더 TimeStamp
	anBrokerCfgCount	: ARRAY[1..3, 1..GVL_MQTT.CONFIG_TOPIC_COUNT] OF UDINT;
	asBrokerCfgTime		: ARRAY[1..3, 1..GVL_MQTT.CONFIG_TOPIC_COUNT] OF STRING(23);
	anPrevCmdCount		: ARRAY[1..3, 1..GVL_MQTT.COMMAND_TOPIC_COUNT] OF UDINT;		// 핸들러가 마지막으로 본 횟수
	anPrevCfgCount		: ARRAY[1..3, 1..GVL_MQTT.CONFIG_TOPIC_COUNT] OF UDINT;
	anCmdRxBroker		: ARRAY[1..GVL_MQTT.COMMAND_TOPIC_COUNT] OF INT;	// 토픽별 마지막으로 받은 브로커 (1 Cloud, 2 Local, 3 Azure)
	anCfgRxBroker		: ARRAY[1..GVL_MQTT.CONFIG_TOPIC_COUNT] OF INT;
	astCmdHeader		: ARRAY[1..GVL_MQTT.COMMAND_TOPIC_COUNT] OF ST_MqttCommandHeader;	// 마지막으로 받은 command 헤더 (Location, SiteID, UserName, TimeStamp, DeviceCount)
	astCfgHeader		: ARRAY[1..GVL_MQTT.CONFIG_TOPIC_COUNT] OF ST_MqttCommandHeader;
	astPcsCommandRx		: ARRAY[0..GVL_PARAM.PCS_COUNT-1] OF ST_MqttCommand_Rx;	// 받은 command/pcs 레코드 사본 (칸 = DeviceIndex - F_MqttDistribute.DEVICE_ID_BASE, 지금 1)
	astBatCommandRx		: ARRAY[0..GVL_PARAM.BMS_COUNT-1] OF ST_MqttCommand_Rx;	// 받은 command/bat 레코드 사본
	astPcsConfigRx		: ARRAY[0..GVL_PARAM.PCS_COUNT-1] OF ST_PcsConfig_Rx;	// 받은 config/pcs 사본
	astBatConfigRx		: ARRAY[0..GVL_PARAM.BMS_COUNT-1] OF ST_BatConfig_Rx;	// 받은 config/bat 사본
	stProtectionConfigRx : ST_ProtectionConfig_Rx;								// 받은 config/protection 사본
	nCmdRxTotal			: UDINT;		// 핸들러가 본 command 수신 누계 (브로커 합)
	nCfgRxTotal			: UDINT;
	sLastRx				: STRING(80);	// 마지막 수신 요약 예) 'Cloud command/pcs 2026-10-21 10:20:00.000'
	pRxHeader			: POINTER TO ST_MqttCommandHeader;
	b					: INT;
	t					: UINT;
END_VAR
VAR CONSTANT
	WAVE_PERIOD		: UDINT := 600;		// 삼각파 주기 (갱신 횟수 = 초)
	PCS_P_MAX		: REAL := 500.0;	// PCS 1대 최대 출력 kW
	BAT_V			: REAL := 740.0;	// DC 전압 V
	AC_V_LL			: REAL := 380.0;	// AC 선간 전압 V
	AC_V_LN			: REAL := 220.0;	// AC 상 전압 V
	SQRT3			: REAL := 1.7320508;
	BROKER_NAME		: ARRAY[1..3] OF STRING(5) := ['Cloud', 'Local', 'Azure'];
END_VAR

IF NOT bEnable THEN
	RETURN;
END_IF

tonUpdate(IN := NOT tonUpdate.Q);
IF NOT (tonUpdate.Q OR NOT bFirstDone) THEN
	RETURN;
END_IF
bFirstDone := TRUE;

(* 공통 값 *)
nTick		:= nTick + 1;
nHeartbeat	:= nTick MOD 100;
fWave		:= ABS(UDINT_TO_REAL(nTick MOD WAVE_PERIOD) / UDINT_TO_REAL(WAVE_PERIOD / 2) - 1.0) * 2.0 - 1.0;	// 1 → -1 → 1
fPcsP		:= PCS_P_MAX * fWave;
fBatSoc		:= 50.0 - 30.0 * fWave;		// 방전(+)할수록 낮음: 20 ~ 80 %
nRacksPerBat := GVL_PARAM.RACKS_PER_BMS;

A_FillPms();
A_FillPcs();
A_FillBat();
A_FillRack();
A_FillPv();
A_FillEss();
A_FillTemp();
A_FillAirConditioner();

ACTION A_FillAirConditioner:
(* 공조기: 냉방·바람 자동 운전, 설정 24 ℃ 근처에서 실내 온도가 오르내림 *)
FOR i := 0 TO GVL_PARAM.AIR_CONDITIONER_COUNT - 1 DO
	fDev := UINT_TO_REAL(i);
	g_stAirConditionerPublish.Devices[i].DeviceIndex		:= UINT_TO_UDINT(i + 1);
	g_stAirConditionerPublish.Devices[i].Status				:= 2#0100;		// b2 운전
	g_stAirConditionerPublish.Devices[i].ModeState			:= 0;			// 0 Cooling
	g_stAirConditionerPublish.Devices[i].WindMode			:= 4;			// 4 Auto
	g_stAirConditionerPublish.Devices[i].ControlTemperature	:= 24.0;		// ℃
	g_stAirConditionerPublish.Devices[i].RoomTemperature	:= 24.0 + 0.2 * fDev + 1.5 * fWave;	// ℃
	g_stAirConditionerPublish.Devices[i].Fault1				:= 0;
END_FOR
END_ACTION

ACTION A_FillBat:
FOR i := 0 TO GVL_PARAM.BMS_COUNT - 1 DO
	fDev := UINT_TO_REAL(i);
	g_stBatPublish.Devices[i].DeviceIndex						:= UINT_TO_UDINT(i + 1);
	g_stBatPublish.Devices[i].Status							:= 0;
	g_stBatPublish.Devices[i].OnlineRackCount					:= UINT_TO_UDINT(nRacksPerBat);
	g_stBatPublish.Devices[i].TotalRackCount					:= UINT_TO_UDINT(nRacksPerBat);
	g_stBatPublish.Devices[i].MaxCellVoltageLocationFromRack	:= 1;
	g_stBatPublish.Devices[i].MaxCellVoltageLocationFromModule	:= 2;
	g_stBatPublish.Devices[i].MaxCellVoltageLocationFromCell	:= 3;
	g_stBatPublish.Devices[i].MinCellVoltageLocationFromRack	:= 4;
	g_stBatPublish.Devices[i].MinCellVoltageLocationFromModule	:= 5;
	g_stBatPublish.Devices[i].MinCellVoltageLocationFromCell	:= 6;
	g_stBatPublish.Devices[i].MaxModuleTempLocationFromRack		:= 7;
	g_stBatPublish.Devices[i].MaxModuleTempLocationFromModule	:= 8;
	g_stBatPublish.Devices[i].MaxModuleTempLocationFromCell		:= 9;
	g_stBatPublish.Devices[i].MinModuleTempLocationFromRack		:= 10;
	g_stBatPublish.Devices[i].MinModuleTempLocationFromModule	:= UINT_TO_UDINT(MIN(UINT#11, GVL_PARAM.MODULES_PER_RACK));
	g_stBatPublish.Devices[i].MinModuleTempLocationFromCell		:= 12;
	g_stBatPublish.Devices[i].Heartbeat							:= nHeartbeat;
	g_stBatPublish.Devices[i].Soc								:= fBatSoc + fDev;			// %
	g_stBatPublish.Devices[i].Soh								:= 98.0 - 0.5 * fDev;		// %
	g_stBatPublish.Devices[i].Eol								:= 80.0;
	g_stBatPublish.Devices[i].DcVoltage							:= BAT_V - 20.0 * fWave;	// 방전할수록 낮음
	g_stBatPublish.Devices[i].DcCurrent							:= fPcsP * 1000.0 / BAT_V;	// A (방전 +)
	g_stBatPublish.Devices[i].ChargeCurrentLimit				:= 800.0;					// A
	g_stBatPublish.Devices[i].DischargeCurrentLimit				:= 800.0;
	g_stBatPublish.Devices[i].ChargePowerLimit					:= 600.0;					// kW
	g_stBatPublish.Devices[i].DischargePowerLimit				:= 600.0;
	g_stBatPublish.Devices[i].MaxCellVoltage					:= 3.35 - 0.05 * fWave;		// V
	g_stBatPublish.Devices[i].MinCellVoltage					:= 3.30 - 0.05 * fWave;
	g_stBatPublish.Devices[i].MaxModuleTemperature				:= 30.0 + 2.0 * ABS(fWave);	// ℃
	g_stBatPublish.Devices[i].MinModuleTemperature				:= 25.0 + ABS(fWave);
	g_stBatPublish.Devices[i].Warning1							:= 0;
	g_stBatPublish.Devices[i].Warning2							:= 0;
	g_stBatPublish.Devices[i].Warning3							:= 0;
	g_stBatPublish.Devices[i].Warning4							:= 0;
	g_stBatPublish.Devices[i].Warning5							:= 0;
	g_stBatPublish.Devices[i].Warning6							:= 0;
	g_stBatPublish.Devices[i].Warning7							:= 0;
	g_stBatPublish.Devices[i].Warning8							:= 0;
	g_stBatPublish.Devices[i].Warning9							:= 0;
	g_stBatPublish.Devices[i].Warning10							:= 0;
	g_stBatPublish.Devices[i].Fault1							:= 0;
	g_stBatPublish.Devices[i].Fault2							:= 0;
	g_stBatPublish.Devices[i].Fault3							:= 0;
	g_stBatPublish.Devices[i].Fault4							:= 0;
	g_stBatPublish.Devices[i].Fault5							:= 0;
	g_stBatPublish.Devices[i].Fault6							:= 0;
	g_stBatPublish.Devices[i].Fault7							:= 0;
	g_stBatPublish.Devices[i].Fault8							:= 0;
	g_stBatPublish.Devices[i].Fault9							:= 0;
	g_stBatPublish.Devices[i].Fault10							:= 0;
END_FOR
END_ACTION

ACTION A_FillEss:
(* ESS 계량: PCS와 같은 방향 (방전 +, 충전 -). 방전량·충전량을 따로 누적 *)
FOR i := 0 TO GVL_PARAM.ESS_COUNT - 1 DO
	fDev := UINT_TO_REAL(i);
	fP := fPcsP * (1.0 - 0.05 * fDev);
	IF fP >= 0.0 THEN
		afEssEnergy[i] := afEssEnergy[i] + fP / 3600.0;
	ELSE
		afEssEnergyRev[i] := afEssEnergyRev[i] - fP / 3600.0;
	END_IF
	g_stEssPublish.Devices[i].EnergyActivePower			:= afEssEnergy[i];		// kWh 방전
	g_stEssPublish.Devices[i].EnergyReactivePower		:= 0.05 * afEssEnergy[i];
	g_stEssPublish.Devices[i].EnergyReverseActivePower	:= afEssEnergyRev[i];	// kWh 충전
	g_stEssPublish.Devices[i].EnergyReverseReactivePower := 0.05 * afEssEnergyRev[i];
	g_stEssPublish.Devices[i].DeviceIndex		:= UINT_TO_UDINT(i + 1);
	g_stEssPublish.Devices[i].Status			:= 1;
	g_stEssPublish.Devices[i].AcActivePower	:= fP;					// kW
	g_stEssPublish.Devices[i].AcReactivePower	:= 0.05 * fP;			// kvar
	g_stEssPublish.Devices[i].AcVoltageR		:= AC_V_LN + fDev;
	g_stEssPublish.Devices[i].AcVoltageS		:= AC_V_LN + fDev + 0.3;
	g_stEssPublish.Devices[i].AcVoltageT		:= AC_V_LN + fDev - 0.3;
	g_stEssPublish.Devices[i].AcCurrentR		:= ABS(fP) * 1000.0 / (3.0 * AC_V_LN);	// A
	g_stEssPublish.Devices[i].AcCurrentS		:= g_stEssPublish.Devices[i].AcCurrentR + 0.3;
	g_stEssPublish.Devices[i].AcCurrentT		:= g_stEssPublish.Devices[i].AcCurrentR - 0.3;
	g_stEssPublish.Devices[i].Frequency		:= 60.0 + 0.02 * fWave;
	g_stEssPublish.Devices[i].PowerFactor		:= 0.99;
	g_stEssPublish.Devices[i].Warning1		:= 0;
	g_stEssPublish.Devices[i].Warning2		:= 0;
	g_stEssPublish.Devices[i].Warning3		:= 0;
	g_stEssPublish.Devices[i].Warning4		:= 0;
	g_stEssPublish.Devices[i].Warning5		:= 0;
	g_stEssPublish.Devices[i].Warning6		:= 0;
	g_stEssPublish.Devices[i].Warning7		:= 0;
	g_stEssPublish.Devices[i].Warning8		:= 0;
	g_stEssPublish.Devices[i].Warning9		:= 0;
	g_stEssPublish.Devices[i].Warning10		:= 0;
	g_stEssPublish.Devices[i].Fault1			:= 0;
	g_stEssPublish.Devices[i].Fault2			:= 0;
	g_stEssPublish.Devices[i].Fault3			:= 0;
	g_stEssPublish.Devices[i].Fault4			:= 0;
	g_stEssPublish.Devices[i].Fault5			:= 0;
	g_stEssPublish.Devices[i].Fault6			:= 0;
	g_stEssPublish.Devices[i].Fault7			:= 0;
	g_stEssPublish.Devices[i].Fault8			:= 0;
	g_stEssPublish.Devices[i].Fault9			:= 0;
	g_stEssPublish.Devices[i].Fault10			:= 0;
END_FOR
END_ACTION

ACTION A_FillPcs:
FOR i := 0 TO GVL_PARAM.PCS_COUNT - 1 DO
	fDev := UINT_TO_REAL(i);
	fP := fPcsP * (1.0 - 0.05 * fDev);		// 장치마다 5 %씩 다르게
	g_stPcsPublish.Devices[i].DeviceIndex			:= UINT_TO_UDINT(i + 1);
	g_stPcsPublish.Devices[i].SystemOperationMode	:= 1;			// 1 모드스케줄
	g_stPcsPublish.Devices[i].OperationMode			:= 1;
	g_stPcsPublish.Devices[i].PMSActivePower		:= fP;			// 지령 kW
	g_stPcsPublish.Devices[i].RemoteMode			:= 1;			// 1 Remote
	g_stPcsPublish.Devices[i].Status				:= 0;
	g_stPcsPublish.Devices[i].AcActivePower			:= fP * 0.99;	// 출력 kW
	g_stPcsPublish.Devices[i].AcReactivePower		:= 0.1 * fP;	// kvar
	g_stPcsPublish.Devices[i].PowerFactor			:= 0.99;
	g_stPcsPublish.Devices[i].Frequency				:= 60.0 + 0.02 * fWave;
	g_stPcsPublish.Devices[i].AcRsVoltage			:= AC_V_LL + fDev;
	g_stPcsPublish.Devices[i].AcStVoltage			:= AC_V_LL + fDev + 0.5;
	g_stPcsPublish.Devices[i].AcTrVoltage			:= AC_V_LL + fDev - 0.5;
	g_stPcsPublish.Devices[i].AcRVoltage			:= AC_V_LN + fDev;
	g_stPcsPublish.Devices[i].AcSVoltage			:= AC_V_LN + fDev + 0.3;
	g_stPcsPublish.Devices[i].AcTVoltage			:= AC_V_LN + fDev - 0.3;
	g_stPcsPublish.Devices[i].AcRCurrent			:= ABS(fP) * 1000.0 / (SQRT3 * AC_V_LL);	// A
	g_stPcsPublish.Devices[i].AcSCurrent			:= g_stPcsPublish.Devices[i].AcRCurrent + 0.5;
	g_stPcsPublish.Devices[i].AcTCurrent			:= g_stPcsPublish.Devices[i].AcRCurrent - 0.5;
	g_stPcsPublish.Devices[i].DcLinkVoltage			:= BAT_V + 10.0;
	g_stPcsPublish.Devices[i].DcVoltage				:= BAT_V;
	g_stPcsPublish.Devices[i].DcCurrent				:= fP * 1000.0 / BAT_V;					// A (방전 +)
	g_stPcsPublish.Devices[i].DcActivePower			:= fP * 1.01;
	g_stPcsPublish.Devices[i].InsulationResistance	:= 2000.0;		// kΩ
	g_stPcsPublish.Devices[i].Temperature1			:= 35.0 + fDev + 3.0 * ABS(fWave);
	g_stPcsPublish.Devices[i].Temperature2			:= 36.0 + fDev + 3.0 * ABS(fWave);
	g_stPcsPublish.Devices[i].Temperature3			:= 37.0 + fDev + 3.0 * ABS(fWave);
	g_stPcsPublish.Devices[i].Temperature4			:= 38.0 + fDev + 3.0 * ABS(fWave);
	g_stPcsPublish.Devices[i].Temperature5			:= 30.0 + fDev;
	g_stPcsPublish.Devices[i].Temperature6			:= 31.0 + fDev;
	g_stPcsPublish.Devices[i].Temperature7			:= 32.0 + fDev;
	g_stPcsPublish.Devices[i].Temperature8			:= 33.0 + fDev;
	g_stPcsPublish.Devices[i].Warning1				:= 0;
	g_stPcsPublish.Devices[i].Warning2				:= 0;
	g_stPcsPublish.Devices[i].Warning3				:= 0;
	g_stPcsPublish.Devices[i].Warning4				:= 0;
	g_stPcsPublish.Devices[i].Warning5				:= 0;
	g_stPcsPublish.Devices[i].Warning6				:= 0;
	g_stPcsPublish.Devices[i].Warning7				:= 0;
	g_stPcsPublish.Devices[i].Warning8				:= 0;
	g_stPcsPublish.Devices[i].Warning9				:= 0;
	g_stPcsPublish.Devices[i].Warning10				:= 0;
	g_stPcsPublish.Devices[i].Fault1				:= 0;
	g_stPcsPublish.Devices[i].Fault2				:= 0;
	g_stPcsPublish.Devices[i].Fault3				:= 0;
	g_stPcsPublish.Devices[i].Fault4				:= 0;
	g_stPcsPublish.Devices[i].Fault5				:= 0;
	g_stPcsPublish.Devices[i].Fault6				:= 0;
	g_stPcsPublish.Devices[i].Fault7				:= 0;
	g_stPcsPublish.Devices[i].Fault8				:= 0;
	g_stPcsPublish.Devices[i].Fault9				:= 0;
	g_stPcsPublish.Devices[i].Fault10				:= 0;
END_FOR
END_ACTION

ACTION A_FillPms:
(* PMS 상태 1건 *)
g_stPmsPublish.Devices[0].DeviceIndex			:= 1;
g_stPmsPublish.Devices[0].Status				:= 1;
g_stPmsPublish.Devices[0].PmsIsAlive			:= 1;			// 1 정상
g_stPmsPublish.Devices[0].CpuUsage				:= 20 + nTick MOD 10;	// %
g_stPmsPublish.Devices[0].CpuTemperature		:= 50;			// ℃
g_stPmsPublish.Devices[0].RemainCycle			:= 80;			// %
g_stPmsPublish.Devices[0].RemainSaveArea		:= 70;			// %
g_stPmsPublish.Devices[0].ProtectModuleCurrent	:= 1.2;
g_stPmsPublish.Devices[0].ProtectModuleVoltage	:= 24.0;
g_stPmsPublish.Devices[0].PmsEvent				:= 0;
g_stPmsPublish.Devices[0].ModuleStatus1			:= 0;
g_stPmsPublish.Devices[0].ModuleStatus2			:= 0;
END_ACTION

ACTION A_FillPv:
(* PV: 낮 발전처럼 100 ~ 300 kW, 누적 발전량은 1 s마다 kW/3600 kWh씩 더함 *)
FOR i := 0 TO GVL_PARAM.PV_COUNT - 1 DO
	fDev := UINT_TO_REAL(i);
	fP := 200.0 + 100.0 * fWave - 10.0 * fDev;
	afPvEnergy[i] := afPvEnergy[i] + fP / 3600.0;
	g_stPvPublish.Devices[i].EnergyActivePower			:= afPvEnergy[i];		// kWh
	g_stPvPublish.Devices[i].EnergyReactivePower		:= 0.05 * afPvEnergy[i];
	g_stPvPublish.Devices[i].EnergyReverseActivePower	:= 0.0;
	g_stPvPublish.Devices[i].EnergyReverseReactivePower	:= 0.0;
	g_stPvPublish.Devices[i].DeviceIndex		:= UINT_TO_UDINT(i + 1);
	g_stPvPublish.Devices[i].Status			:= 1;
	g_stPvPublish.Devices[i].AcActivePower	:= fP;					// kW
	g_stPvPublish.Devices[i].AcReactivePower	:= 0.05 * fP;			// kvar
	g_stPvPublish.Devices[i].AcVoltageR		:= AC_V_LN + fDev;
	g_stPvPublish.Devices[i].AcVoltageS		:= AC_V_LN + fDev + 0.3;
	g_stPvPublish.Devices[i].AcVoltageT		:= AC_V_LN + fDev - 0.3;
	g_stPvPublish.Devices[i].AcCurrentR		:= ABS(fP) * 1000.0 / (3.0 * AC_V_LN);	// A
	g_stPvPublish.Devices[i].AcCurrentS		:= g_stPvPublish.Devices[i].AcCurrentR + 0.3;
	g_stPvPublish.Devices[i].AcCurrentT		:= g_stPvPublish.Devices[i].AcCurrentR - 0.3;
	g_stPvPublish.Devices[i].Frequency		:= 60.0 + 0.02 * fWave;
	g_stPvPublish.Devices[i].PowerFactor		:= 0.99;
	g_stPvPublish.Devices[i].Warning1		:= 0;
	g_stPvPublish.Devices[i].Warning2		:= 0;
	g_stPvPublish.Devices[i].Warning3		:= 0;
	g_stPvPublish.Devices[i].Warning4		:= 0;
	g_stPvPublish.Devices[i].Warning5		:= 0;
	g_stPvPublish.Devices[i].Warning6		:= 0;
	g_stPvPublish.Devices[i].Warning7		:= 0;
	g_stPvPublish.Devices[i].Warning8		:= 0;
	g_stPvPublish.Devices[i].Warning9		:= 0;
	g_stPvPublish.Devices[i].Warning10		:= 0;
	g_stPvPublish.Devices[i].Fault1			:= 0;
	g_stPvPublish.Devices[i].Fault2			:= 0;
	g_stPvPublish.Devices[i].Fault3			:= 0;
	g_stPvPublish.Devices[i].Fault4			:= 0;
	g_stPvPublish.Devices[i].Fault5			:= 0;
	g_stPvPublish.Devices[i].Fault6			:= 0;
	g_stPvPublish.Devices[i].Fault7			:= 0;
	g_stPvPublish.Devices[i].Fault8			:= 0;
	g_stPvPublish.Devices[i].Fault9			:= 0;
	g_stPvPublish.Devices[i].Fault10			:= 0;
END_FOR
END_ACTION

ACTION A_FillRack:
(* 번호·BatID·ModuleCount는 PRG_PublishDeviceNo에서 채움. 여기서는 시험 측정값만 생성 *)
FOR i := 0 TO GVL_PARAM.RACK_COUNT - 1 DO
	fDev := UINT_TO_REAL(i MOD 10);			// 10개 주기로 조금씩 다르게
	g_stRackPublish.Devices[i].Status			:= 1;
	g_stRackPublish.Devices[i].Soc				:= fBatSoc + 0.2 * fDev;		// %
	g_stRackPublish.Devices[i].Soh				:= 98.0 - 0.1 * fDev;
	g_stRackPublish.Devices[i].DcVoltage		:= BAT_V - 20.0 * fWave + 0.5 * fDev;
	g_stRackPublish.Devices[i].DcCurrent		:= fPcsP * 1000.0 / BAT_V / UINT_TO_REAL(nRacksPerBat);	// A
	g_stRackPublish.Devices[i].ChargeCurrentLimit		:= 100.0;
	g_stRackPublish.Devices[i].DischargeCurrentLimit	:= 100.0;
	g_stRackPublish.Devices[i].ChargePowerLimit			:= 70.0;
	g_stRackPublish.Devices[i].DischargePowerLimit		:= 70.0;
	g_stRackPublish.Devices[i].AvgCellVoltage	:= 3.32 - 0.05 * fWave;
	g_stRackPublish.Devices[i].MaxCellVoltage	:= 3.35 - 0.05 * fWave;
	g_stRackPublish.Devices[i].MinCellVoltage	:= 3.29 - 0.05 * fWave;
	g_stRackPublish.Devices[i].AvgModuleTemp	:= 27.0 + 0.1 * fDev;
	g_stRackPublish.Devices[i].MaxModuleTemp	:= 30.0 + 0.1 * fDev;
	g_stRackPublish.Devices[i].MinModuleTemp	:= 24.0 + 0.1 * fDev;
	g_stRackPublish.Devices[i].MaxCellVoltageLocationFromModule	:= (i MOD GVL_PARAM.MODULES_PER_RACK) + 1;
	g_stRackPublish.Devices[i].MaxCellVoltageLocationFromCell	:= (i MOD 16) + 1;
	g_stRackPublish.Devices[i].MinCellVoltageLocationFromModule	:= ((i + 3) MOD GVL_PARAM.MODULES_PER_RACK) + 1;
	g_stRackPublish.Devices[i].MinCellVoltageLocationFromCell	:= ((i + 5) MOD 16) + 1;
	g_stRackPublish.Devices[i].MaxModuleTempLocationFromModule	:= ((i + 1) MOD GVL_PARAM.MODULES_PER_RACK) + 1;
	g_stRackPublish.Devices[i].MaxModuleTempLocationFromCell	:= ((i + 7) MOD 16) + 1;
	g_stRackPublish.Devices[i].MinModuleTempLocationFromModule	:= ((i + 4) MOD GVL_PARAM.MODULES_PER_RACK) + 1;
	g_stRackPublish.Devices[i].MinModuleTempLocationFromCell	:= ((i + 9) MOD 16) + 1;
	g_stRackPublish.Devices[i].Warning1			:= 0;
	g_stRackPublish.Devices[i].Warning2			:= 0;
	g_stRackPublish.Devices[i].Warning3			:= 0;
	g_stRackPublish.Devices[i].Warning4			:= 0;
	g_stRackPublish.Devices[i].Warning5			:= 0;
	g_stRackPublish.Devices[i].Warning6			:= 0;
	g_stRackPublish.Devices[i].Warning7			:= 0;
	g_stRackPublish.Devices[i].Warning8			:= 0;
	g_stRackPublish.Devices[i].Warning9			:= 0;
	g_stRackPublish.Devices[i].Warning10		:= 0;
	g_stRackPublish.Devices[i].Fault1			:= 0;
	g_stRackPublish.Devices[i].Fault2			:= 0;
	g_stRackPublish.Devices[i].Fault3			:= 0;
	g_stRackPublish.Devices[i].Fault4			:= 0;
	g_stRackPublish.Devices[i].Fault5			:= 0;
	g_stRackPublish.Devices[i].Fault6			:= 0;
	g_stRackPublish.Devices[i].Fault7			:= 0;
	g_stRackPublish.Devices[i].Fault8			:= 0;
	g_stRackPublish.Devices[i].Fault9			:= 0;
	g_stRackPublish.Devices[i].Fault10			:= 0;
END_FOR
END_ACTION

ACTION A_FillTemp:
(* 온도·습도 센서. location 1 PCS실, 2 BAT실, 3 UPS실, 4 FC 컨테이너실, 5 외부 *)
FOR i := 0 TO GVL_PARAM.TEMP_COUNT - 1 DO
	fDev := UINT_TO_REAL(i);
	g_stTempPublish.Devices[i].DeviceIndex	:= UINT_TO_UDINT(i + 1);
	g_stTempPublish.Devices[i].status		:= 1;
	g_stTempPublish.Devices[i].location		:= UINT_TO_UDINT(i MOD 5) + 1;
	g_stTempPublish.Devices[i].temperature	:= 24.0 + fDev + 2.0 * fWave;	// ℃
	g_stTempPublish.Devices[i].humidity		:= 45.0 + 2.0 * fDev + 5.0 * fWave;	// %
END_FOR
END_ACTION

ACTION A_HandleRx:
(* 수신 시험 핸들러: 새로 받은 command·config를 브로커·토픽별로 기록하고 레코드 사본을 남김
   PRG_Mqtt가 FB_MqttMain(구독·분배) 다음, FB_EmsCommand(CommandType 지움) 앞에서 PRG_MqttTestData.A_HandleRx()로 부름 *)

(* 1. 브로커별 수신 횟수·시각 (1 Cloud, 2 Local, 3 Azure) *)
FOR t := 1 TO GVL_MQTT.COMMAND_TOPIC_COUNT DO
	anBrokerCmdCount[1, t] := PRG_Mqtt.fbMqttMain.fbCloudSub.q_anCmdRxCount[t];	asBrokerCmdTime[1, t] := PRG_Mqtt.fbMqttMain.fbCloudSub.q_asCmdRxTime[t];
	anBrokerCmdCount[2, t] := PRG_Mqtt.fbMqttMain.fbLocalSub.q_anCmdRxCount[t];	asBrokerCmdTime[2, t] := PRG_Mqtt.fbMqttMain.fbLocalSub.q_asCmdRxTime[t];
	anBrokerCmdCount[3, t] := PRG_Mqtt.fbMqttMain.fbAzureSub.q_anCmdRxCount[t];	asBrokerCmdTime[3, t] := PRG_Mqtt.fbMqttMain.fbAzureSub.q_asCmdRxTime[t];
END_FOR
FOR t := 1 TO GVL_MQTT.CONFIG_TOPIC_COUNT DO
	anBrokerCfgCount[1, t] := PRG_Mqtt.fbMqttMain.fbCloudSub.q_anCfgRxCount[t];	asBrokerCfgTime[1, t] := PRG_Mqtt.fbMqttMain.fbCloudSub.q_asCfgRxTime[t];
	anBrokerCfgCount[2, t] := PRG_Mqtt.fbMqttMain.fbLocalSub.q_anCfgRxCount[t];	asBrokerCfgTime[2, t] := PRG_Mqtt.fbMqttMain.fbLocalSub.q_asCfgRxTime[t];
	anBrokerCfgCount[3, t] := PRG_Mqtt.fbMqttMain.fbAzureSub.q_anCfgRxCount[t];	asBrokerCfgTime[3, t] := PRG_Mqtt.fbMqttMain.fbAzureSub.q_asCfgRxTime[t];
END_FOR

(* 2. command: 횟수가 바뀐 브로커·토픽 = 새 메시지 (헤더 TimeStamp가 바뀐 것) *)
FOR b := 1 TO 3 DO
	FOR t := 1 TO GVL_MQTT.COMMAND_TOPIC_COUNT DO
		IF anBrokerCmdCount[b, t] <> anPrevCmdCount[b, t] THEN
			anPrevCmdCount[b, t] := anBrokerCmdCount[b, t];
			anCmdRxBroker[t] := b;
			nCmdRxTotal := nCmdRxTotal + 1;
			pRxHeader := PRG_Mqtt.fbMqttMain.astSubCommandTable[t].pRxBuffer;
			IF pRxHeader <> 0 THEN
				astCmdHeader[t] := pRxHeader^;
			END_IF
			IF t = 1 THEN
				astPcsCommandRx := g_astPcsCommand;		// FB_EmsCommand가 지우기 전 사본
			ELSE
				astBatCommandRx := g_astBatCommand;
			END_IF
			sLastRx := CONCAT(CONCAT(BROKER_NAME[b], ' command/'), CONCAT(PRG_Mqtt.fbMqttMain.astSubCommandTable[t].sTopic, CONCAT(' ', asBrokerCmdTime[b, t])));
		END_IF
	END_FOR
END_FOR

(* 3. config *)
FOR b := 1 TO 3 DO
	FOR t := 1 TO GVL_MQTT.CONFIG_TOPIC_COUNT DO
		IF anBrokerCfgCount[b, t] <> anPrevCfgCount[b, t] THEN
			anPrevCfgCount[b, t] := anBrokerCfgCount[b, t];
			anCfgRxBroker[t] := b;
			nCfgRxTotal := nCfgRxTotal + 1;
			pRxHeader := PRG_Mqtt.fbMqttMain.astSubConfigTable[t].pRxBuffer;
			IF pRxHeader <> 0 THEN
				astCfgHeader[t] := pRxHeader^;
			END_IF
			CASE t OF
				1:	astPcsConfigRx := g_astPcsConfig;
				2:	astBatConfigRx := g_astBatConfig;
				3:	stProtectionConfigRx := g_stProtectionConfig;
			END_CASE
			sLastRx := CONCAT(CONCAT(BROKER_NAME[b], ' config/'), CONCAT(PRG_Mqtt.fbMqttMain.astSubConfigTable[t].sTopic, CONCAT(' ', asBrokerCfgTime[b, t])));
		END_IF
	END_FOR
END_FOR
END_ACTION

END_PROGRAM

// ---- 99_Test/PRG_TestLogger.TcPOU
PROGRAM PRG_TestLogger		// 로거(MQTT 로거 토픽, 지금 pms_log) 시험 (GVL_SITE.TEST_MODE일 때 PRG_Mqtt가 부름): 이벤트 로거에 등록된 이벤트를 찾아 보내고, 브로커 대신 큐에서 패킷을 꺼내 확인. 브로커 접속 없이 됨
// 버튼은 온라인에서 TRUE로 쓰면 1회 하고 FALSE로 돌아감 (bAlarm만 켜 두는 스위치)
// 등록된 이벤트 (시작할 때 자동으로 찾음. 이벤트를 추가·삭제·변경해도 이 프로그램은 고치지 않음)
//   클래스 4개(TC_EVENT_CLASSES: PmsSystem·PmsProt·PmsOutput·PmsSeq) × 번호 1..SCAN_ID_MAX를 이벤트 로거에 문구 요청 → 문구가 오면 등록된 이벤트
//   bScanDone 뒤 nFound(찾은 수), astReg[n]: 이름(클래스 번호)·문구 틀(인자 자리 #0#~#5#)·인자 수·고정 글자·남는 글자(95 − 고정)·확인 필요
//   확인 필요(bCheck, nCheck) = 고정 글자 FIXED_MAX(50) 초과 또는 인자 하나당 남는 글자(nPerArg)가 ARG_MIN(10)자 미만 → 문구 틀을 줄이거나 실제 인자 길이를 확인 (PMS_STD.md 7장 "로그 문구 길이")
// 보내기 (인자 자리에는 문구 틀에 적힌 그대로 {0}, {1} … 를 넣음 → Error List·EMS에 문구 틀 모양 그대로 보임)
//   bSendAll 찾은 것 전부 (스캔마다 SEND_PER_SCAN건) → bAllDone 뒤 bAllOk (다 받음 + 잘린 수 = 예상 nExpectTrunc + 문구 오류 0)
//   bSendOne nSendNo번 한 건, bSendNext nSendNo번 보내고 다음 번호로 (wsSendName, wsLastSent)
//   문구가 실제 로그와 같게 Error List·EMS에 나감 (심각도는 모두 Info: 원래 심각도는 PLC에서 읽을 수 없음)
// 로거 경로 시험 (시험 이벤트 PmsSystem.LoggerTest "로거 시험: {0}{1}")
//   bAlarm 켜면 알람 발생 "로거 시험: 알람", 끄면 해소 "[해소] 로거 시험: 알람" (등록된 이벤트 보내기는 메시지만 보내서 알람 경로는 여기서만 시험)
//   bSendLong 127자 메시지 → 99자 + '…'로 잘리고 PRG_Mqtt.fbMqttMain.fbLogger.q_nTruncated 1 증가
// 받은 로그: awsAllRx·asAllRxTime (큐에서 꺼낸 전체 로그, ALL_KEEP칸을 돌려 씀, 마지막 칸 = nAllRxLast)
VAR
	(* 로거 경로 시험 *)
	bAlarm			: BOOL;			// TRUE = 알람 발생, FALSE = 해소
	bSendLong		: BOOL;			// 127자 메시지 1건
	(* 등록된 이벤트 (자동으로 찾음) *)
	bScanDone		: BOOL;			// 찾기 끝 (시작 뒤 약 5 s)
	wsScanStep		: WSTRING(40);	// 찾는 중인 클래스·번호, 끝나면 찾은 수
	nFound			: UINT;			// 찾은 이벤트 수
	nCheck			: UINT;			// 확인 필요 수
	nScanMiss		: UINT;			// 없는 번호(오류·빈 문구·시간 초과)로 건너뛴 수
	nScanOverflow	: UINT;			// REG_MAX를 넘어 못 담은 수 (0이어야 함)
	astReg			: ARRAY[1..REG_MAX] OF ST_LoggerTestReg;
	(* 보내기 *)
	bSendAll		: BOOL;			// 찾은 것 전부
	bSendOne		: BOOL;			// nSendNo번 한 건
	bSendNext		: BOOL;			// nSendNo번 한 건 보내고 다음 번호로
	nSendNo			: UINT := 1;	// 1..nFound
	wsSendName		: WSTRING(31);	// nSendNo번 이벤트 (클래스 번호)
	wsLastSent		: WSTRING(31);	// 마지막으로 보낸 이벤트
	bAllBusy		: BOOL;			// 보내는 중 또는 받기를 기다리는 중
	bAllDone		: BOOL;
	bAllOk			: BOOL;			// 다 받음 + 잘린 수 = 예상 + 문구 오류 0
	nAllRx			: UDINT;		// 보낸 뒤 받은 로그 수 (실제 로그가 끼면 더 많을 수 있음)
	nAllTrunc		: UDINT;		// 그동안 100자를 넘어 잘린 수
	nExpectTrunc	: UDINT;		// 잘릴 것으로 계산한 수 (고정 + 인자 수 × 3자 > 100. 보통 0)
	nAllTextErr		: UDINT;
	(* 받은 로그 (큐에서 꺼낸 순서) *)
	nAllRxCount		: UDINT;
	nAllRxLast		: UINT;
	awsAllRx		: ARRAY[1..ALL_KEEP] OF WSTRING(100);
	asAllRxTime		: ARRAY[1..ALL_KEEP] OF STRING(23);
	(* 내부 *)
	bInit			: BOOL;
	nNext			: UDINT;		// 이 시험이 큐에서 꺼낼 다음 번호 (브로커와 따로)
	stPacket		: ST_LoggerPublish_V1;
	fbMsg			: FB_LogMsg;
	fbAlarm			: FB_LogAlarm;
	asArg			: ARRAY[1..6] OF WSTRING(63);
	asAlarmArg		: ARRAY[1..6] OF WSTRING(63) := ["알람", 5("")];
	aClassGuid		: ARRAY[1..CLASS_COUNT] OF GUID;
	awsClassName	: ARRAY[1..CLASS_COUNT] OF WSTRING(15);
	fbScanText		: FB_RequestEventText;
	fbScanArgs		: FB_TcMessage;		// 문구 틀 분석용 인자(#0#~#5#)만 담음. 보내지 않음
	tonScan			: TON := (PT := T#2S);
	nScanState		: UINT;			// 0 준비, 1 요청, 2 받기, 3 끝
	nScanClass		: UINT;
	nScanId			: UDINT;
	{attribute 'TcEncoding' := 'UTF-8'}
	sScanText		: STRING(511);
	wsText			: WSTRING(255);
	wsWork			: WSTRING(255);
	wsMark			: WSTRING(5);
	wsTrail			: WSTRING(8);	// 문구 끝에 덧붙은 인자 표시 " (#n#)"
	bTrail			: BOOL;
	bArgUsed		: BOOL;
	nArgs			: UINT;
	nFixed			: UINT;
	nPos			: INT;
	afbReg			: ARRAY[1..REG_MAX] OF FB_LogMsg;
	asFill			: ARRAY[1..6] OF WSTRING(63);	// 보낼 인자: {0} … {5} (A_InitScan)
	nRegIdx			: UINT;
	nSendIdx		: UINT;
	nAllStartRx		: UDINT;
	nAllTruncBefore	: UDINT;
	nAllTextErrBefore : UDINT;
	tonAll			: TON := (PT := T#5S);
	i				: UINT;
	k				: UINT;
END_VAR
VAR CONSTANT
	CLASS_COUNT		: UINT := 4;		// 찾는 이벤트 클래스 수 (A_InitScan, 로거 리스너 필터와 같은 클래스)
	SCAN_ID_MAX		: UDINT := 64;		// 클래스마다 찾아보는 번호 (1..64)
	REG_MAX			: UINT := 64;		// 담을 수 있는 이벤트 수
	TEXT_RULE		: UINT := 95;		// 로그 문구 규칙 (PMS_STD.md 7장)
	FIXED_MAX		: UINT := 50;		// 문구 틀 고정 글자 권장 한도
	ARG_MIN			: UINT := 10;		// 판정: 인자 하나당 남는 글자가 이보다 적으면 확인 필요
	SEND_PER_SCAN	: UINT := 32;		// bSendAll이 한 스캔에 보내는 수 (로거 큐 GVL_MQTT.LOGGER_QUEUE 64칸 안)
	ALL_KEEP		: UINT := 70;
END_VAR

IF NOT bInit THEN
	bInit := TRUE;
	nNext := PRG_Mqtt.fbMqttMain.fbLogger.q_nReceived + 1;		// 시작 전 로그는 건너뜀
	A_InitScan();
END_IF

fbMsg(i_stEntry := TC_EVENTS.PmsSystem.LoggerTest);
IF bSendLong THEN
	bSendLong := FALSE;
	A_SendLong();
END_IF
fbAlarm(i_stEntry := TC_EVENTS.PmsSystem.LoggerTest, i_bActive := bAlarm, i_nArgs := 2, i_asArg := asAlarmArg);

A_Scan();
A_Send();
A_Receive();

ACTION A_AddReg:
// 찾은 이벤트 한 칸: 문구 틀(wsText, 인자 자리 #n#)을 분석해 인자 수·고정 글자·확인 필요를 정하고, 보낼 FB를 이 이벤트로 정함
IF nFound >= REG_MAX THEN
	nScanOverflow := nScanOverflow + 1;
	RETURN;
END_IF
nFound := nFound + 1;

// TwinCAT은 문구 자리보다 많이 넘긴 인자를 문구 끝에 " (값)"으로 덧붙인다 (요청할 때 6개를 넘기므로).
// 끝에서부터 " (#5#)", " (#4#)" … 을 떼어 내고 남은 것이 문구 틀이다.
// 한계: 문구 틀이 맨 끝에서 " ({n})"으로 끝나면 덧붙은 것과 구분하지 못함 (2026-10-28 기준 그런 문구 없음)
bTrail := TRUE;
FOR k := 0 TO 5 DO
	IF bTrail THEN
		wsTrail := WCONCAT(WCONCAT(" (#", TO_WSTRING(5 - k)), "#)");
		nPos := WLEN(wsText) - WLEN(wsTrail) + 1;
		IF nPos >= 1 AND_THEN WMID(wsText, WLEN(wsTrail), nPos) = wsTrail THEN
			wsText := WLEFT(wsText, nPos - 1);
		ELSE
			bTrail := FALSE;
		END_IF
	END_IF
END_FOR

astReg[nFound].stEntry.uuidEventClass	:= aClassGuid[nScanClass];
astReg[nFound].stEntry.nEventId			:= nScanId;
astReg[nFound].stEntry.eSeverity		:= TcEventSeverity.Info;
astReg[nFound].wsName					:= WCONCAT(WCONCAT(awsClassName[nScanClass], " "), TO_WSTRING(nScanId));
astReg[nFound].wsTemplate				:= wsText;

// 인자 자리 표시(#n#, 인자가 안 들어갔으면 {n})를 지운 길이 = 고정 글자. 인자 수 = 쓰인 가장 큰 번호 + 1
wsWork	:= wsText;
nArgs	:= 0;
FOR i := 0 TO 5 DO
	bArgUsed := FALSE;
	wsMark := WCONCAT(WCONCAT("#", TO_WSTRING(i)), "#");
	A_StripMark();
	wsMark := WCONCAT(WCONCAT("{", TO_WSTRING(i)), "}");
	A_StripMark();
	IF bArgUsed THEN
		nArgs := i + 1;
	END_IF
END_FOR
nFixed := INT_TO_UINT(WLEN(wsWork));
astReg[nFound].nArgs	:= nArgs;
astReg[nFound].nFixed	:= nFixed;
astReg[nFound].nFree	:= UINT_TO_INT(TEXT_RULE) - UINT_TO_INT(nFixed);
IF nArgs > 0 AND nFixed < TEXT_RULE THEN
	astReg[nFound].nPerArg := (TEXT_RULE - nFixed) / nArgs;
ELSIF nArgs > 0 THEN
	astReg[nFound].nPerArg := 0;
ELSE
	astReg[nFound].nPerArg := TEXT_RULE - MIN(nFixed, TEXT_RULE);
END_IF
astReg[nFound].bCheck	:= nFixed > FIXED_MAX OR astReg[nFound].nPerArg < ARG_MIN;
IF astReg[nFound].bCheck THEN
	nCheck := nCheck + 1;
END_IF
afbReg[nFound].i_stEntry := astReg[nFound].stEntry;		// FB_LogMsg는 처음 보낼 때 이 이벤트로 만들어짐
END_ACTION

ACTION A_InitScan:
// 찾을 클래스 (로거 리스너 필터와 같은 4개. 새 이벤트 클래스를 만들면 여기와 CLASS_COUNT에도 더함)
aClassGuid[1] := TC_EVENT_CLASSES.PmsSystem;	awsClassName[1] := "PmsSystem";
aClassGuid[2] := TC_EVENT_CLASSES.PmsProt;		awsClassName[2] := "PmsProt";
aClassGuid[3] := TC_EVENT_CLASSES.PmsOutput;	awsClassName[3] := "PmsOutput";
aClassGuid[4] := TC_EVENT_CLASSES.PmsSeq;		awsClassName[4] := "PmsSeq";

// 문구 틀 분석용 인자: 인자 자리마다 표시 #0#~#5# (이 메시지는 만들기만 하고 보내지 않음)
fbScanArgs.CreateEx(stEventEntry := TC_EVENTS.PmsSystem.LoggerTest, ipSourceInfo := 0);
fbScanArgs.ipArguments.Clear();
FOR i := 0 TO 5 DO
	wsMark := WCONCAT(WCONCAT("#", TO_WSTRING(i)), "#");
	fbScanArgs.ipArguments.AddWString(wsMark);
END_FOR

// 보낼 인자: 문구 틀에 적힌 그대로 {0} … {5}
FOR i := 1 TO 6 DO
	asFill[i] := WCONCAT(WCONCAT("{", TO_WSTRING(i - 1)), "}");
END_FOR

nScanClass	:= 1;
nScanId		:= 1;
nScanState	:= 1;
END_ACTION

ACTION A_Receive:
// 브로커 대신 큐에서 꺼냄 (스캔마다 준비된 것 전부)
FOR i := 1 TO 40 DO
	IF NOT PRG_Mqtt.fbMqttMain.fbLogger.M_GetPacket(i_nSiteId := GVL_SITE.MQTT_SET.nSiteId, iq_nNext := nNext, iq_stPacket := stPacket) THEN
		EXIT;
	END_IF
	nNext := nNext + 1;
	nAllRxCount				:= nAllRxCount + 1;
	nAllRxLast				:= UDINT_TO_UINT(((nAllRxCount - 1) MOD ALL_KEEP) + 1);
	awsAllRx[nAllRxLast]	:= stPacket.Contents;
	asAllRxTime[nAllRxLast]	:= stPacket.Header.TimeStamp;
END_FOR
END_ACTION

ACTION A_Scan:
// 등록된 이벤트 찾기: 클래스·번호마다 문구를 요청해 문구가 오면 등록된 것. 한 번에 하나씩 (시작 뒤 약 5 s)
CASE nScanState OF
	1:	// 요청
		wsScanStep := WCONCAT(WCONCAT(awsClassName[nScanClass], " "), TO_WSTRING(nScanId));
		fbScanText.Clear();
		fbScanText.Request(eventClass := aClassGuid[nScanClass], nEventId := nScanId,
						nLangId := GVL_MQTT.LOGGER_LANG_ID, ipArgs := fbScanArgs.ipArguments);
		tonScan(IN := FALSE);
		nScanState := 2;

	2:	// 받기: 오류·빈 문구·시간 초과 = 없는 번호
		tonScan(IN := TRUE);
		IF fbScanText.bError OR tonScan.Q THEN
			nScanMiss := nScanMiss + 1;
			A_ScanNext();
		ELSIF NOT fbScanText.bBusy THEN
			sScanText := '';
			fbScanText.GetString(sScanText, SIZEOF(sScanText));
			wsText := F_Utf8ToWstring(i_pSrc := ADR(sScanText), i_nSrcSize := SIZEOF(sScanText));
			// 없는 번호: 빈 문구, 또는 런타임이 돌려주는 "EventText not found…" (4024.17은 오류 대신 이 문구)
			IF wsText = "" OR WFIND(wsText, "EventText not found") = 1 THEN
				nScanMiss := nScanMiss + 1;
			ELSE
				A_AddReg();
			END_IF
			A_ScanNext();
		END_IF
END_CASE
END_ACTION

ACTION A_ScanNext:
// 다음 번호, 클래스 끝이면 다음 클래스, 모두 끝이면 찾기 끝
tonScan(IN := FALSE);
nScanId := nScanId + 1;
IF nScanId > SCAN_ID_MAX THEN
	nScanId		:= 1;
	nScanClass	:= nScanClass + 1;
END_IF
IF nScanClass > CLASS_COUNT THEN
	nScanState	:= 3;
	bScanDone	:= TRUE;
	wsScanStep	:= WCONCAT(TO_WSTRING(nFound), "종 찾음");
ELSE
	nScanState := 1;
END_IF
END_ACTION

ACTION A_Send:
// 보내기 버튼 (누르면 1회 하고 FALSE로). 찾기가 끝나야 보냄
IF nSendNo < 1 OR nSendNo > MAX(nFound, 1) THEN
	nSendNo := 1;
END_IF
IF nFound > 0 THEN
	wsSendName := astReg[nSendNo].wsName;
END_IF
IF NOT bScanDone OR nFound = 0 THEN
	bSendAll	:= FALSE;
	bSendOne	:= FALSE;
	bSendNext	:= FALSE;
	RETURN;
END_IF

// 인자는 {0} … {5} 그대로 (A_InitScan에서 한 번 채움)

IF bSendOne THEN
	bSendOne := FALSE;
	nRegIdx := nSendNo;
	A_SendReg();
END_IF
IF bSendNext THEN
	bSendNext := FALSE;
	nRegIdx := nSendNo;
	A_SendReg();
	nSendNo := (nSendNo MOD nFound) + 1;
END_IF

IF bSendAll THEN
	bSendAll			:= FALSE;
	nSendIdx			:= 1;
	nAllStartRx			:= nAllRxCount;
	nAllTruncBefore		:= PRG_Mqtt.fbMqttMain.fbLogger.q_nTruncated;
	nAllTextErrBefore	:= PRG_Mqtt.fbMqttMain.fbLogger.q_nTextError;
	nExpectTrunc		:= 0;
	FOR i := 1 TO nFound DO
		IF astReg[i].nFixed + astReg[i].nArgs * 3 > INT_TO_UINT(GVL_MQTT.LOGGER_TEXT_MAX) THEN
			nExpectTrunc := nExpectTrunc + 1;
		END_IF
	END_FOR
	bAllBusy	:= TRUE;
	bAllDone	:= FALSE;
	bAllOk		:= FALSE;
	tonAll(IN := FALSE);
END_IF

IF bAllBusy THEN
	// 스캔마다 SEND_PER_SCAN건씩 (로거 큐를 넘지 않게)
	k := 0;
	WHILE nSendIdx <= nFound AND k < SEND_PER_SCAN DO
		nRegIdx := nSendIdx;
		A_SendReg();
		nSendIdx	:= nSendIdx + 1;
		k			:= k + 1;
	END_WHILE
	// 다 보낸 뒤: 다 받음 + 잘린 수가 예상과 같음 + 문구 오류 없음
	IF nSendIdx > nFound THEN
		tonAll(IN := TRUE);
		nAllRx := nAllRxCount - nAllStartRx;
		IF nAllRx >= nFound OR tonAll.Q THEN
			bAllBusy	:= FALSE;
			bAllDone	:= TRUE;
			nAllTrunc	:= PRG_Mqtt.fbMqttMain.fbLogger.q_nTruncated - nAllTruncBefore;
			nAllTextErr	:= PRG_Mqtt.fbMqttMain.fbLogger.q_nTextError - nAllTextErrBefore;
			bAllOk		:= nAllRx >= nFound AND nAllTrunc = nExpectTrunc AND nAllTextErr = 0;
			tonAll(IN := FALSE);
		END_IF
	END_IF
END_IF
END_ACTION

ACTION A_SendLong:
// 고정 7자 + 인자 60자 + 60자 = 127자 → 99자 + '…'로 잘려야 함
asArg[1] := "012345678901234567890123456789012345678901234567890123456789";
asArg[2] := asArg[1];
fbMsg.M_SendEvent(2, asArg);
END_ACTION

ACTION A_SendReg:
// 찾은 이벤트 nRegIdx 한 건 (인자 수만큼 {0} … 를 넣음)
afbReg[nRegIdx].M_SendEvent(astReg[nRegIdx].nArgs, asFill);
wsLastSent := astReg[nRegIdx].wsName;
END_ACTION

ACTION A_StripMark:
// wsWork에서 wsMark를 모두 지움. 하나라도 있으면 bArgUsed
nPos := WFIND(wsWork, wsMark);
WHILE nPos > 0 DO
	wsWork		:= WDELETE(wsWork, WLEN(wsMark), nPos);
	bArgUsed	:= TRUE;
	nPos		:= WFIND(wsWork, wsMark);
END_WHILE
END_ACTION

END_PROGRAM

// ---- 10_Core/70_Diag/FB_LogMsg.TcPOU
FUNCTION_BLOCK FB_LogMsg		// 메시지 한 종류: M_SendEvent 할 때마다 1회 기록
VAR_INPUT
	i_stEntry		: TcEventEntry;
END_VAR
VAR
	_fbMsg			: FB_TcMessage;
	_bInit			: BOOL;
END_VAR

IF NOT _bInit THEN
	_fbMsg.CreateEx(stEventEntry := i_stEntry, ipSourceInfo := 0);
	_bInit := TRUE;
END_IF

METHOD M_SendEvent
VAR_INPUT
	i_nArgs		: UINT;
	i_asArg		: ARRAY[1..6] OF WSTRING(63);
END_VAR
VAR
	k			: UINT;
END_VAR
IF NOT _bInit THEN
	_fbMsg.CreateEx(stEventEntry := i_stEntry, ipSourceInfo := 0);
	_bInit := TRUE;
END_IF
_fbMsg.ipArguments.Clear();
FOR k := 1 TO MIN(i_nArgs, 6) DO
	_fbMsg.ipArguments.AddWString(i_asArg[k]);
END_FOR
_fbMsg.Send(0);
END_METHOD

END_FUNCTION_BLOCK

// ---- 10_Core/70_Diag/FB_LogAlarm.TcPOU
FUNCTION_BLOCK FB_LogAlarm		// 알람 하나: 켜질 때 발생 1회, 꺼질 때 해소 1회. 인자는 발생할 때 한 번 넣음
VAR_INPUT
	i_stEntry		: TcEventEntry;		// 등록한 이벤트 (TC_EVENTS.클래스.이벤트). 심각도는 처음 만들 때 값
	i_bActive		: BOOL;
	i_nArgs			: UINT;				// 인자 수 (0~6)
	i_asArg			: ARRAY[1..6] OF WSTRING(63);
END_VAR
VAR_OUTPUT
	q_bRaised		: BOOL;				// 지금 발생 중 (호출 전에 이 값과 i_bActive가 다를 때만 인자를 만들면 됨)
END_VAR
VAR
	_fbAlarm		: FB_TcAlarm;
	_bInit			: BOOL;
END_VAR
VAR_TEMP
	k				: UINT;
END_VAR

IF NOT _bInit THEN
	_fbAlarm.CreateEx(stEventEntry := i_stEntry, bWithConfirmation := FALSE, ipSourceInfo := 0);
	_bInit := TRUE;
END_IF

IF i_bActive AND NOT q_bRaised THEN
	_fbAlarm.ipArguments.Clear();
	FOR k := 1 TO MIN(i_nArgs, 6) DO
		_fbAlarm.ipArguments.AddWString(i_asArg[k]);
	END_FOR
	_fbAlarm.Raise(0);
	q_bRaised := TRUE;
ELSIF NOT i_bActive AND q_bRaised THEN
	_fbAlarm.Clear(0, FALSE);
	q_bRaised := FALSE;
END_IF

END_FUNCTION_BLOCK

// ---- 90_Project/MAIN.TcPOU
PROGRAM MAIN
VAR
	fbSnapshot		: FB_Snapshot;
	fbMeasure		: FB_Measure;
	fbProtection	: FB_Protection;
	fbBatGroup		: FB_BatGroup;
	fbUnitAvail	: FB_UnitAvail;
	fbEquipLimits	: FB_EquipmentLimits;
	fbGroupView		: FB_GroupView;
	fbUnitView		: FB_UnitView;		// 유닛(PCS)마다 요약 (유닛 단위 제어 모드 관리자가 봄)
	fbSources		: FB_SourceHub;
	fbModeSwitch	: FB_ModeSwitch;
	fbStateArb		: FB_StateArbiter;
	fbSelect		: FB_Select;
	fbAutoGate		: FB_Gate;
	fbManualGate	: FB_Gate;
	fbOutputReady	: FB_OutputReady;
	fbLimitEval		: FB_LimitEval;
	fbManualShape	: FB_ShapePath := (i_bManual := TRUE);
	fbAutoShape		: FB_ShapePath := (i_bManual := FALSE);
	fbDistributor	: FB_Distributor;
	fbSequencer		: FB_Sequencer;
	fbPermitEval	: FB_PermitEval;	// 기동 조건 모듈 평가
	fbGroupState	: FB_GroupState;	// 그룹 상태 요약
	fbDispatcher	: FB_Dispatcher;
	fbAuxOutput		: FB_AuxOutput;
	fbOutputDiag	: FB_OutputDiag;
	fbEventLog		: FB_EventLog;
	fbAlive			: FB_AliveRecorder;
	fbPersistSave	: FB_PersistSave;
	fbConfigCheck	: FB_ConfigCheck;
	fbSettingGuard	: FB_SettingGuard;	// 운전 중 바꾸는 설정 값 지키기
	fbModuleList	: FB_ModuleList;
	fbReport		: FB_Report;
	fbClock			: FB_LocalClock;	// 현지 시각 (제어 모드 시간표)
	afZeroGrp		: ARRAY[1..GVL_PARAM.GROUP_COUNT] OF REAL;		// Manual 성형의 '다른 경로 몫' (없음 = 0)
	bTestReset		: BOOL;		// 시험 리셋 (TEST_MODE AND GVL_TEST.g_bTestReset): 모든 PCS·BMS 고장 리셋 + 유지 DO 풀기
	bClearHoldDo	: BOOL;		// 유지 DO 풀기: 지금은 지령원 PCS 리셋 요청·시험 리셋과 같은 신호 (DO 작업 때 따로 정함)
	stUpsConfigReceived : ST_IfUpsConfigRx; // coherent received snapshot. 주기적·펄스 값만 fbUpsConfigApply가 적용
	fbUpsConfigApply : ARRAY[1..GVL_PARAM.UPS_COUNT] OF FB_UpsConfigApply; // EMS 설정 → UPS 쓰기
	nUpsConfigReadSeq : UDINT;
	stUpsConfigCandidate : ST_IfUpsConfigRx;
	nUpsCmdReadSeq : UDINT; // GVL_IF.g_nUpsCmdSeq 읽은 값
	astUpsCmdCandidate : ARRAY[1..GVL_PARAM.UPS_COUNT] OF ST_IfUpsCmd;
	astUpsCmdReceived : ARRAY[1..GVL_PARAM.UPS_COUNT] OF ST_IfUpsCmd; // 일관되게 읽은 UPS 명령
	fbUpsCommand : ARRAY[1..GVL_PARAM.UPS_COUNT] OF FB_UpsCommand; // EMS UPS 명령 → UPS 명령 레지스터 (명세 WR-UPS-01)
	bUpsConfigOk : BOOL;
	_nReportPcs : UINT; // action loop variable, not VAR_TEMP
// 통신 시험 중 충방전 알고리즘 선언 중지 (2026-11-02)
// afbUpsCharge : ARRAY[1..GVL_PARAM.UPS_COUNT] OF FB_UpsChargeSequence;
// afbUpsTemp : ARRAY[1..GVL_PARAM.UPS_COUNT] OF FB_UpsTemperatureCharge;
// astUpsChargeSet : ARRAY[1..GVL_PARAM.UPS_COUNT] OF ST_UpsChargeSet; // 미확정 값은 0
// aeUpsChargeMode : ARRAY[1..GVL_PARAM.UPS_COUNT] OF E_UpsChargeMode;
// abUpsChargeEnable : ARRAY[1..GVL_PARAM.UPS_COUNT] OF BOOL;
// abUpsChargeCancel : ARRAY[1..GVL_PARAM.UPS_COUNT] OF BOOL;
// abUpsChargeReset : ARRAY[1..GVL_PARAM.UPS_COUNT] OF BOOL;
// abUpsTempEnable : ARRAY[1..GVL_PARAM.UPS_COUNT] OF BOOL;
// astUpsChargeFeedback : ARRAY[1..GVL_PARAM.UPS_COUNT] OF ST_UpsChargeFeedback;
// astUpsTempFeedback : ARRAY[1..GVL_PARAM.UPS_COUNT] OF ST_UpsChargeFeedback;
 fbRptBat : ARRAY[1..GVL_PARAM.BMS_COUNT] OF FB_RptEsolutionBat; // 배터리 보고 매핑
 _nReportBat : UINT; // 배터리 보고 번호
 _nReportRack : UINT; // 랙 보고 번호
 _nReportModule : UINT; // 모듈 보고 번호
 fbRptUps : ARRAY[1..GVL_PARAM.UPS_COUNT] OF FB_RptSebangUps; // UPS 보고 매핑
 fbRptImd : ARRAY[1..GVL_PARAM.IMD_COUNT] OF FB_RptLsImd1000; // IMD 보고 매핑 (토픽 imd)
 _nReportImd : UINT; // IMD 보고 번호
 fbRptTemp : ARRAY[1..GVL_PARAM.TEMP_COUNT] OF FB_RptTempHum; // 온습도 보고 매핑 (토픽 temperature_sensor)
 fbBmsRack : ARRAY[1..GVL_PARAM.BMS_COUNT] OF FB_BmsRackCommand; // 랙 컨택터 개별 제어 (EMS CommandType 11·12)
 abBmsRackAcc : ARRAY[1..GVL_PARAM.BMS_COUNT] OF BOOL; // 지난 스캔 랙 쓰기 요청을 드라이버가 받음
 aeBmsRackRes : ARRAY[1..GVL_PARAM.BMS_COUNT] OF E_UpsResult; // 지난 스캔 드라이버 결과
 fbBmsCtl : ARRAY[1..GVL_PARAM.BMS_COUNT] OF FB_BmsContactorCommand; // 컨택터 하나씩 제어 (EMS CommandType 5~10) [2026-11-13]
 abBmsCtlAcc : ARRAY[1..GVL_PARAM.BMS_COUNT] OF BOOL; // 지난 스캔 컨택터 쓰기 요청을 드라이버가 받음
 aeBmsCtlRes : ARRAY[1..GVL_PARAM.BMS_COUNT] OF E_UpsResult; // 지난 스캔 드라이버 결과
 fbUpsSafety : ARRAY[1..GVL_PARAM.UPS_COUNT] OF FB_UpsSafetyStage; // 사고·고장 단계 판정 (UPS n ↔ BMS n). 표시만, 장비에 쓰지 않음
 // BMS 쓰기 시험 (시뮬레이터 전용). 값을 넣고 nBmsTestCmd를 쓰면 1회 실행 후 0으로 돌아감
 // 1 랙 비트(wBmsTestValue), 2 충전 접촉기, 3 방전 접촉기, 4 시스템 접촉기(bBmsTestOn), 5 비상차단, 6 리셋, 7 주기적 방전 시작, 8 방전 취소
 nBmsTestCmd : UINT;
 wBmsTestValue : WORD := 16#00FF; // 랙 비트. b0 = 랙 1 (랙 8개)
 bBmsTestOn : BOOL; // 접촉기 On/Off
 eBmsTestResult : E_UpsResult; // 마지막 접수 결과
 stBmsTestCmd : ST_BatCmd;
 nBmsTestSeq : UDINT := 16#80000000; // 코어 명령 번호와 겹치지 않게
 _nReportUps : UINT; // UPS 보고 번호
	awsUpsConfigError : ARRAY[1..GVL_PARAM.UPS_COUNT] OF WSTRING(63);
	bWriteEnable	: BOOL;		// 장비 쓰기 허가 (설정 오류 없음 AND 주 PLC AND DEVICE_WRITE). 디스패처·보조 출력·시퀀서가 씀
	stEmsCopy		: ST_IfEmsCmd;	// MQTT 명령 칸의 마지막 일관된 복사본
	nEmsSeq			: UDINT;
	fbEmsCfg		: FB_EmsConfigApply;	// EMS config(pcs·bat) → 운영 설정 [9-21 수정 2026-11-04: 추가]
	stEmsCfgCopy	: ST_IfEmsCfg;		// MQTT config 칸의 마지막 복사본
	nEmsCfgSeq		: UDINT;
	bEmsCfgOk		: BOOL;
	stEmsOut		: ST_SourceOutput;	// EMS 지령원 출력 (지난 스캔). 속성 결과는 칸을 바로 못 읽어 한 번 담음
	(* [16번 수정 2026-11-09: 추가] A_PassEmsCmd: PCS 지령 → 스탠다드 스케줄 유닛 칸 (액션이라 VAR에 둠) *)
	nCmU			: UINT;
	nCmK			: UINT;
	nCmPcs			: UINT;
	fCmPcsRated		: REAL;
	fbBrokerWatch	: FB_BrokerWatch;	// MQTT 브로커 끊김 감시 [9번 수정 2026-11-09: 추가]
END_VAR
VAR_TEMP
	i			: UINT;
END_VAR

(* ===== 0. 가상 장비 연결 (시험 모드에서만. 현장은 GVL_SITE.TEST_MODE = FALSE) ===== *)
IF GVL_SITE.TEST_MODE THEN
	PRG_SimLink();
	PRG_TestCtrlMode();	// 제어 모드 자동 시험 (따로 둔 인스턴스만 씀. 결과 PRG_TestCtrlMode.fbTally)
	PRG_TestSchedLive();	// 스케줄 모드 실제 경로 시험 (bStart := TRUE로 시작할 때만 동작)
	PRG_TestPeakLive();	// 피크컷·통합 모드 실제 경로 시험 (bStart := TRUE로 시작할 때만 동작)
	PRG_TestUnitMode();	// 유닛 단위 제어 모드 자동 시험 (따로 둔 인스턴스만 씀. 결과 PRG_TestUnitMode.fbTally). [16번 수정 2026-11-09: 현장 PCS별 실경로 시험 PRG_TestUnitLive는 없앰]
	PRG_TestStdLive();	// 스탠다드 스케줄 모드 실제 경로 시험 (EMS 명령 → 모드 → 코어 고르기. bStart := TRUE로 시작)
END_IF

(* ===== 현지 시각 (A_PassModuleSet이 제어 모드 관리자에 넘김) ===== *)
fbClock();

(* ===== 모듈 설정 넘기기: GVL_PERSIST.g_stModuleSet 칸 → 모듈 i_stSet (A_PassModuleSet, 현장 모듈마다 한 줄) ===== *)
A_PassEmsCfg();		// [9-21 수정 2026-11-04: 추가] EMS config → GVL_PERSIST 설정 (모듈 설정 넘기기 앞: 같은 스캔에 모듈·설정 보호가 새 값을 봄)
A_PassModuleSet();
A_PassEmsCmd();
// Raw config mailbox only. Do not drive charge modes from this received structure.
// UPS 명령 칸 (MqttTask → PlcTask): 번호가 짝수이고 복사 전후가 같을 때만 받음
nUpsCmdReadSeq:=GVL_IF.g_nUpsCmdSeq;
IF (nUpsCmdReadSeq AND 1)=0 THEN
 astUpsCmdCandidate:=GVL_IF.g_astUpsCmd;
 IF nUpsCmdReadSeq=GVL_IF.g_nUpsCmdSeq THEN astUpsCmdReceived:=astUpsCmdCandidate; END_IF
END_IF
nUpsConfigReadSeq:=GVL_IF.g_nUpsConfigSeq;
IF (nUpsConfigReadSeq AND 1)=0 THEN
 stUpsConfigCandidate:=GVL_IF.g_stUpsConfigRx;
 IF nUpsConfigReadSeq=GVL_IF.g_nUpsConfigSeq THEN stUpsConfigReceived:=stUpsConfigCandidate; END_IF
END_IF

(* ===== 등록된 모듈 목록: 모듈 ID 점검·로그 이름 찾기는 이 목록만 봄 (새 등록 배열은 FB_ModuleList에만 추가) ===== *)
fbModuleList(	iq_aipPcs	:= GVL_SITE.g_aipPcs,
				iq_aipBms	:= GVL_SITE.g_aipBms,
				iq_aipMeter	:= GVL_SITE.g_aipMeter,
				iq_aipAux	:= GVL_SITE.g_aipAux,
				iq_aipSource	:= GVL_SITE.g_aipSource,
				iq_aipLimit	:= GVL_SITE.g_aipLimit,
				iq_aipPermit	:= GVL_SITE.g_aipPermit,
				iq_aipComp	:= GVL_SITE.g_aipComp,
				iq_aipRule	:= GVL_SITE.g_aipRule,
				iq_aipResp	:= GVL_SITE.g_aipResp,
				iq_aipOutput	:= GVL_SITE.g_aipOutput,
				iq_aipUnitRule	:= GVL_SITE.g_aipUnitRule,
				iq_aipBatRule	:= GVL_SITE.g_aipBatRule,
				iq_aipSelPolicy	:= GVL_SITE.g_aipSelectPolicy,
				iq_aipDistPolicy	:= GVL_SITE.g_aipDistPolicy,
				iq_ipAutoGate	:= GVL_SITE.g_ipAutoGate,
				iq_ipManualGate	:= GVL_SITE.g_ipManualGate,
				iq_astUnitCfg	:= GVL_SITE.UNIT_CFG);

(* ===== 운전 중 바꾸는 설정 지키기: 잘못된 값은 마지막 정상값으로 되돌림 (GVL_PERSIST에 다시 씀). 모듈 설정을 되돌렸으면 다시 넘김 ===== *)
fbSettingGuard(	i_pModuleSet	:= ADR(GVL_PERSIST.g_stModuleSet),
				i_nModuleSetSize	:= SIZEOF(GVL_PERSIST.g_stModuleSet),
				iq_stCmdFilter	:= GVL_PERSIST.g_stCmdFilter,
				iq_stManualCmdSet	:= GVL_PERSIST.g_stManualCmdSet,
				iq_stSeqSet		:= GVL_PERSIST.g_stSeqSet,
				iq_astGroupSet	:= GVL_PERSIST.g_astGroupSet,	// [결함 13 수정 2026-11-04: 추가]
				iq_aipModule	:= fbModuleList.q_aipModule,
				iq_astOutputCfg	:= GVL_PERSIST.g_astOutputCfg,
				iq_astRuleCfg	:= GVL_PERSIST.g_astRuleCfg,
				iq_astSourceReg	:= GVL_PERSIST.g_astSourceReg,
				iq_astLimitReg	:= GVL_PERSIST.g_astLimitReg,
				iq_astPermitReg	:= GVL_PERSIST.g_astPermitReg,
				iq_astCompReg	:= GVL_PERSIST.g_astCompReg,
				iq_astUnitRuleReg	:= GVL_PERSIST.g_astUnitRuleReg,
				iq_astBatRuleReg	:= GVL_PERSIST.g_astBatRuleReg,
				iq_aipLimit		:= GVL_SITE.g_aipLimit,
				iq_aipPermit	:= GVL_SITE.g_aipPermit,
				iq_aipComp		:= GVL_SITE.g_aipComp,
				iq_aipRule		:= GVL_SITE.g_aipRule);
IF fbSettingGuard.q_bRestored THEN
	A_PassModuleSet();
END_IF

(* ===== EMS config echo: 설정 보호 뒤 실제 설정 → GVL_IF (MQTT가 config echo로 발행) [9-21 수정 2026-11-04: 추가] ===== *)
fbEmsCfg.M_BuildEcho(	iq_stSocLimit	:= GVL_PERSIST.g_stModuleSet.stSocLimit,
						iq_stUnitLimit	:= GVL_PERSIST.g_stModuleSet.stUnitLimit);
GVL_IF.g_nCfgEchoSeq	:= GVL_IF.g_nCfgEchoSeq + 1;
GVL_IF.g_stEmsCfgEcho	:= fbEmsCfg.q_stEcho;
GVL_IF.g_nCfgEchoSeq	:= GVL_IF.g_nCfgEchoSeq + 1;

(* ===== 설정 점검 (매 스캔): 오류면 장비 쓰기 전부 차단 (디스패처·보조 출력·시퀀서 명령) ===== *)
fbConfigCheck(	iq_astUnitCfg	:= GVL_SITE.UNIT_CFG,
				iq_astBmsCfg	:= GVL_SITE.BMS_CFG,
				iq_astGroupCfg	:= GVL_SITE.GROUP_CFG,
				iq_astPointCfg	:= GVL_SITE.POINT_CFG,
				i_bModuleSetTooBig	:= fbSettingGuard.q_bModuleSetTooBig,
				i_bSetNoGood	:= fbSettingGuard.q_bNoGood,
				i_sSetNoGood	:= fbSettingGuard.q_sNoGood,
				i_stRedSet		:= GVL_SITE.RED_SET,
				i_eRedRole		:= GVL_IF.g_eRedRole,
				iq_aipModule	:= fbModuleList.q_aipModule,
				iq_aipCtrlMode	:= GVL_SITE.g_aipCtrlMode1,	// [2번 수정 2026-11-09: 제어 모드 ID 점검]
				iq_abUnitInstalled	:= fbModuleList.q_abUnitInstalled);

(* ===== 1. 읽기 · 스냅샷 · 계측 ===== *)
// UPS is a separate device type; no PCS power/set-state mapping is used.
bUpsConfigOk:=TRUE;
FOR i:=1 TO GVL_PARAM.UPS_COUNT DO
 awsUpsConfigError[i]:="";
 IF GVL_SITE.g_aipUps[i]<>0 THEN
  awsUpsConfigError[i]:=GVL_SITE.g_aipUps[i].M_CheckSet();
  IF awsUpsConfigError[i]<>"" THEN bUpsConfigOk:=FALSE; END_IF
 END_IF
 IF GVL_SITE.UPS_BMS[i]<1 OR GVL_SITE.UPS_BMS[i]>GVL_PARAM.BMS_COUNT THEN bUpsConfigOk:=FALSE; END_IF
END_FOR
bWriteEnable := fbConfigCheck.q_bConfigOk AND GVL_IF.g_bRedWrite AND GVL_SITE.DEVICE_WRITE AND bUpsConfigOk;
GVL_SITE.g_fbUps1.i_bWritePermit:=bWriteEnable;
GVL_SITE.g_fbBms1.i_bWritePermit:=bWriteEnable;
FOR i:=1 TO GVL_PARAM.UPS_COUNT DO
 IF GVL_SITE.g_aipUps[i]<>0 THEN GVL_SITE.g_aipUps[i].M_Cycle(); END_IF
END_FOR
fbUpsConfigApply[1](i_bEnable:=bWriteEnable AND GVL_PARAM.UPS_CONTROL_ENABLED, i_nRxCount:=stUpsConfigReceived.nRxCount,
 i_stConfig:=stUpsConfigReceived.astConfig[0], i_stState:=GVL_SITE.g_fbUps1.q_stState, i_stRaw:=GVL_SITE.g_fbUps1.q_stRaw, i_ipUps:=GVL_SITE.g_aipUps[1],
 i_bUpsFault:=fbRptUps[1].q_stUps.Status.2, iq_stDesired:=GVL_PERSIST.g_astUpsDesired[1]);
FOR i:=1 TO GVL_PARAM.UPS_COUNT DO
 fbUpsCommand[i](i_stCmd:=astUpsCmdReceived[i], i_bEnable:=bWriteEnable AND GVL_PARAM.UPS_CONTROL_ENABLED,
  i_stUps:=fbRptUps[i].q_stUps, i_bUpsValid:=fbRptUps[i].q_bValid, i_ipUps:=GVL_SITE.g_aipUps[i],
  iq_stDesired:=GVL_PERSIST.g_astUpsDesired[i]);
END_FOR

FOR i := 1 TO GVL_PARAM.PCS_COUNT DO
	IF GVL_SITE.g_aipPcs[i] <> 0 THEN GVL_SITE.g_aipPcs[i].M_Cycle(); END_IF
END_FOR
FOR i := 1 TO GVL_PARAM.BMS_COUNT DO
	IF GVL_SITE.g_aipBms[i] <> 0 THEN GVL_SITE.g_aipBms[i].M_Cycle(); END_IF
END_FOR
FOR i := 1 TO GVL_PARAM.METER_COUNT DO
	IF GVL_SITE.g_aipMeter[i] <> 0 THEN GVL_SITE.g_aipMeter[i].M_Cycle(); END_IF
END_FOR
FOR i := 1 TO GVL_PARAM.AUX_COUNT DO
	IF GVL_SITE.g_aipAux[i] <> 0 THEN GVL_SITE.g_aipAux[i].M_Cycle(); END_IF
END_FOR
fbSnapshot(	iq_aipPcs		:= GVL_SITE.g_aipPcs,
			iq_aipBms		:= GVL_SITE.g_aipBms,
			iq_aipMeter		:= GVL_SITE.g_aipMeter,
			iq_astUnitCfg	:= GVL_SITE.UNIT_CFG);

fbMeasure(	i_bTestMode		:= GVL_SITE.TEST_MODE,
			iq_astMeter		:= fbSnapshot.q_astMeter,
			iq_astPointCfg	:= GVL_SITE.POINT_CFG,
			iq_astGroupCfg	:= GVL_SITE.GROUP_CFG,
			iq_astVirtual	:= GVL_TEST.g_astVirtual);

(* ===== 2. 운전 모드 · 보호 판단 · 유닛 가용 ===== *)
// 고장 리셋은 장비 명령일 뿐 (시퀀서가 지령원 요청을 장비별로 봄). 유지 DO 풀기는 따로 (지령원 요청은 지난 스캔 값: 지령원이 뒤에 돌기 때문)
bTestReset		:= GVL_SITE.TEST_MODE AND GVL_TEST.g_bTestReset;
bClearHoldDo	:= bTestReset OR fbSources.q_bReset;

// 운전 모드: 요청(GVL_PERSIST.g_aeOpMode) → 전환 시퀀스 → 실제 모드. 아래는 모두 실제 모드를 씀 (동작은 그대로, 보호가 실제 모드를 써서 앞에서 부름)
(* ===== MQTT 브로커 끊김 → 운전 모드 요청을 모두 Manual로 (끊김마다 한 번, Active PLC만) [9번 수정 2026-11-09: 추가] ===== *)
fbBrokerWatch(	i_stSet			:= GVL_PERSIST.g_stBrokerWatch,
				i_abUse			:= GVL_IF.g_abBrokerUse,
				i_abConnected	:= GVL_IF.g_abBrokerConn,
				i_bActive		:= GVL_IF.g_bRedActive);
IF fbBrokerWatch.q_bToManual THEN
	FOR i := 1 TO GVL_PARAM.UNIT_COUNT DO
		GVL_PERSIST.g_aeOpMode[i] := E_OpMode.Manual;
	END_FOR
END_IF

fbModeSwitch(	i_stSet			:= GVL_SITE.MODE_SET,
				i_fDonePct		:= GVL_PERSIST.g_stSeqSet.stPcs.fStopDonePct,
				iq_aeModeReq	:= GVL_PERSIST.g_aeOpMode,
				iq_astUnit		:= fbSnapshot.q_astUnit,
				iq_astUnitCfg	:= GVL_SITE.UNIT_CFG,
				iq_astUnitProt	:= fbProtection.q_astUnitProt);	// 지난 스캔 보호 결과: ToManual이면 요청 모드를 Manual로 바꿈

fbProtection(	iq_astUnit		:= fbSnapshot.q_astUnit,
				iq_astBms		:= fbSnapshot.q_astBms,
				iq_astPcc		:= fbMeasure.q_astPcc,
				iq_astUnitCfg	:= GVL_SITE.UNIT_CFG,
				iq_astBmsCfg	:= GVL_SITE.BMS_CFG,
				iq_astRuleCfg	:= GVL_PERSIST.g_astRuleCfg,
				iq_abUnitInstalled	:= fbModuleList.q_abUnitInstalled,
				iq_abBmsInstalled	:= fbModuleList.q_abBmsInstalled,
				iq_aeOpMode		:= fbModeSwitch.q_aeOpMode,
				iq_aipRule		:= GVL_SITE.g_aipRule,
				iq_aipResp		:= GVL_SITE.g_aipResp);

fbBatGroup(		iq_astBms		:= fbSnapshot.q_astBms,
				iq_astBmsCfg	:= GVL_SITE.BMS_CFG,
				iq_astBmsProt	:= fbProtection.q_astBmsProt,
				iq_abBmsInstalled	:= fbModuleList.q_abBmsInstalled);

fbUnitAvail(	iq_astUnit		:= fbSnapshot.q_astUnit,
				iq_astUnitCfg	:= GVL_SITE.UNIT_CFG,
				iq_astUnitProt	:= fbProtection.q_astUnitProt,
				iq_astBatGroup	:= fbBatGroup.q_astBatGroup,
				iq_abUnitInstalled	:= fbModuleList.q_abUnitInstalled);

// 설비 한도: 유닛(정격 × Derate ∩ 유닛 제한 모듈), 배터리 버스(BMS 한도 ∩ 버스 제한 모듈), 그룹 설비 범위. 성형·분배가 같이 씀
fbEquipLimits(	iq_astUnitCfg	:= GVL_SITE.UNIT_CFG,
				iq_astUnit	:= fbSnapshot.q_astUnit,
				iq_astAvail	:= fbUnitAvail.q_astAvail,
				iq_astUnitProt	:= fbProtection.q_astUnitProt,
				iq_aeOpMode	:= fbModeSwitch.q_aeOpMode,
				iq_astBatGroup	:= fbBatGroup.q_astBatGroup,
				iq_astUnitRuleReg	:= GVL_PERSIST.g_astUnitRuleReg,
				iq_astBatRuleReg	:= GVL_PERSIST.g_astBatRuleReg,
				iq_aipUnitRule	:= GVL_SITE.g_aipUnitRule,
				iq_aipBatRule	:= GVL_SITE.g_aipBatRule);

(* ===== 3. 요청 (지령원) ===== *)
fbGroupView(	iq_astPcc		:= fbMeasure.q_astPcc,
				iq_astUnit		:= fbSnapshot.q_astUnit,
				iq_astAvail		:= fbUnitAvail.q_astAvail,
				iq_astUnitCfg	:= GVL_SITE.UNIT_CFG,
				iq_astBatGroup	:= fbBatGroup.q_astBatGroup,
				iq_aeGroupState	:= fbGroupState.q_aeGroupState,	// 지난 스캔
				iq_astGroupEnv	:= fbEquipLimits.q_astGroupEnv);

// 유닛(PCS)마다 요약: 유닛 단위 제어 모드 관리자가 봄 (A_PassModuleSet이 주소를 넘김. 지령원보다 먼저)
fbUnitView(		iq_astView		:= fbGroupView.q_astView,
				iq_astUnit		:= fbSnapshot.q_astUnit,
				iq_astAvail		:= fbUnitAvail.q_astAvail,
				iq_astUnitCfg	:= GVL_SITE.UNIT_CFG,
				iq_astUnitEnv	:= fbEquipLimits.q_astUnitEnv,
				iq_astBatGroup	:= fbBatGroup.q_astBatGroup,
				iq_astBatEnv	:= fbEquipLimits.q_astBatEnv);

fbSources(		iq_aipSource	:= GVL_SITE.g_aipSource,
				iq_astReg		:= GVL_PERSIST.g_astSourceReg,
				iq_astView		:= fbGroupView.q_astView);

(* ===== 4. [제어 그룹마다] 중재 · 성형 (Auto 경로·Manual 경로가 같은 단계) ===== *)

// 상태 요청: 이번 스캔 조건 준비 → 요청 후보 → 접수 검사 → 접수된 것만 이번 스캔 요청 (명령은 6.의 시퀀서 본체가 한 번 보냄)
// 기동 조건 모듈: 그룹마다 한 번 평가 (기다리는 중 표시는 시퀀서 지난 스캔)
fbPermitEval(	iq_astView		:= fbGroupView.q_astView,
				iq_astPermitReg	:= GVL_PERSIST.g_astPermitReg,
				iq_abWaitPermit	:= fbSequencer.q_abWaitPermit,
				iq_aipPermit	:= GVL_SITE.g_aipPermit);

// 장비 쓰기 허가: 설정 오류 없음 + 이 PLC가 Active이고 쓰기 대기가 지남 (PRG_Redundancy) + 장비 쓰기 스위치 (GVL_SITE.DEVICE_WRITE). 대기 PLC는 계산만 하고 장비에 쓰지 않음 (이중화를 안 쓰면 항상 허가)
// 시퀀서도 쓰기 불가를 알고 명령을 만들지 않으며 기동 요청은 거부함 (접수 검사 전에 정해야 해서 여기서 계산)
// Write permission is computed immediately before the device cycle above.

fbSequencer.M_Prepare(	i_bCmdEnable	:= fbConfigCheck.q_bConfigOk,
						i_bWriteEnable	:= bWriteEnable,
						iq_aeStartMode	:= GVL_SITE.START_MODE,
						iq_astUnit		:= fbSnapshot.q_astUnit,
						iq_astAvail		:= fbUnitAvail.q_astAvail,
						iq_astUnitCfg	:= GVL_SITE.UNIT_CFG,
						iq_astBatGroup	:= fbBatGroup.q_astBatGroup,
						iq_abPermit		:= fbPermitEval.q_abPermit,
						iq_abUnitInstalled	:= fbModuleList.q_abUnitInstalled);	// [결함 6 수정 2026-11-03: 추가. 원래 iq_abPermit 뒤에서 끝남]

fbStateArb(		iq_astSrcOut	:= fbSources.q_astOut,
				iq_anSrcModule	:= fbSources.q_anModule,
				iq_astReg		:= GVL_PERSIST.g_astSourceReg,
				iq_aeOpMode		:= fbModeSwitch.q_aeOpMode,
				iq_astUnitCfg	:= GVL_SITE.UNIT_CFG,
				iq_astUnitProt	:= fbProtection.q_astUnitProt,
				iq_abSwitching	:= fbModeSwitch.q_abSwitching);

fbSequencer.M_CheckRequest(	iq_abCand		:= fbStateArb.q_abCand,
							iq_aeCand		:= fbStateArb.q_aeCand);

fbStateArb.M_CommitRequest(iq_abAccept := fbSequencer.q_abAccept);

fbSelect(		iq_aipSelPolicy	:= GVL_SITE.g_aipSelectPolicy,
				iq_astSrcOut	:= fbSources.q_astOut,
				iq_anSrcModule	:= fbSources.q_anModule,
				iq_astReg		:= GVL_PERSIST.g_astSourceReg,
				iq_aeOpMode		:= fbModeSwitch.q_aeOpMode,
				iq_astUnitCfg	:= GVL_SITE.UNIT_CFG,
				iq_astGroupSet	:= GVL_PERSIST.g_astGroupSet,
				iq_astView		:= fbGroupView.q_astView,
				iq_stFilter		:= GVL_PERSIST.g_stCmdFilter);

// 지령 거르기: Auto 경로 (지금은 그대로 통과) / Manual 경로 (방향 반대 무시, 새 지령 표시, Run 뒤 새 지령 대기)
fbAutoGate(		i_ePath			:= E_OpMode.Auto,
				i_ipGate		:= GVL_SITE.g_ipAutoGate,
				iq_astUnitP		:= fbSelect.q_astAutoUnitP,
				iq_astUnitQ		:= fbSelect.q_astAutoUnitQ,
				iq_astGrpP		:= fbSelect.q_astAutoGrpP,
				iq_astGrpQ		:= fbSelect.q_astAutoGrpQ,
				iq_aeOpMode		:= fbModeSwitch.q_aeOpMode,
				iq_astUnit		:= fbSnapshot.q_astUnit,
				iq_astUnitCfg	:= GVL_SITE.UNIT_CFG);

fbManualGate(	i_ePath			:= E_OpMode.Manual,
				i_ipGate			:= GVL_SITE.g_ipManualGate,
				i_stManualCmdSet	:= GVL_PERSIST.g_stManualCmdSet,
				iq_astUnitP			:= fbSelect.q_astManualUnitP,
				iq_astUnitQ			:= fbSelect.q_astManualUnitQ,
				iq_astGrpP			:= fbSelect.q_astManualGrpP,
				iq_astGrpQ			:= fbSelect.q_astManualGrpQ,
				iq_aeOpMode			:= fbModeSwitch.q_aeOpMode,
				iq_astUnit			:= fbSnapshot.q_astUnit,
				iq_astUnitCfg	:= GVL_SITE.UNIT_CFG);

// 출력 가능 유닛: 가용 + 장비 활성(Run·대기) + 정지 진행 중 아님 + 전환 아님 + 새 지령 대기 아님. 성형·분배·디스패처가 이 결과만 씀
fbOutputReady(	iq_astAvail	:= fbUnitAvail.q_astAvail,
				iq_astUnit	:= fbSnapshot.q_astUnit,
				iq_abStopping	:= fbSequencer.q_abStopping,	// 지난 스캔
				iq_abSwitching	:= fbModeSwitch.q_abSwitching,
				iq_abManualWaitNewCmd	:= fbManualGate.q_abWaitNewCmd);

// 제한·보정 모듈: 그룹마다 한 번 평가 (두 경로가 같은 결과를 씀)
fbLimitEval(	iq_astView		:= fbGroupView.q_astView,
				iq_astLimitReg	:= GVL_PERSIST.g_astLimitReg,
				iq_astCompReg	:= GVL_PERSIST.g_astCompReg,
				iq_aipLimit		:= GVL_SITE.g_aipLimit,
				iq_aipComp		:= GVL_SITE.g_aipComp);

// 성형: Manual 경로 먼저 → Auto 경로 (같은 FB. Auto는 접속점 제한을 Manual 몫까지 합쳐 봄)
fbManualShape(	iq_astView			:= fbGroupView.q_astView,
				iq_astGroupSet		:= GVL_PERSIST.g_astGroupSet,
				iq_astManualPolicy	:= GVL_PERSIST.g_astManualPolicy,
				iq_astUnitCfg		:= GVL_SITE.UNIT_CFG,
				iq_aeOpMode			:= fbModeSwitch.q_aeOpMode,
				iq_abOutputReady	:= fbOutputReady.q_abReady,
				iq_astUnitP			:= fbManualGate.q_astUnitP,
				iq_astUnitQ			:= fbManualGate.q_astUnitQ,
				iq_astGrpP			:= fbManualGate.q_astGrpP,
				iq_astGrpQ			:= fbManualGate.q_astGrpQ,
				iq_astGrpPLim		:= fbSelect.q_astManualGrpPLim,
				iq_astGrpQLim		:= fbSelect.q_astManualGrpQLim,
				iq_afOtherGrpP		:= afZeroGrp,
				iq_afOtherGrpQ		:= afZeroGrp,
				iq_aabLimOn			:= fbLimitEval.q_aabOn,
				iq_aastLim			:= fbLimitEval.q_aastLim,
				iq_aaeBasis			:= fbLimitEval.q_aaeBasis,
				iq_aanLimModule		:= fbLimitEval.q_aanModule,
				iq_abPccManual		:= fbLimitEval.q_abPccManual,
				iq_abResume			:= fbLimitEval.q_abResume,
				iq_afPComp			:= fbLimitEval.q_afPComp,
				iq_afQComp	:= fbLimitEval.q_afQComp,
				iq_astGroupEnv	:= fbEquipLimits.q_astGroupEnv);

fbAutoShape(	iq_astView			:= fbGroupView.q_astView,
				iq_astGroupSet		:= GVL_PERSIST.g_astGroupSet,
				iq_astManualPolicy	:= GVL_PERSIST.g_astManualPolicy,
				iq_astUnitCfg		:= GVL_SITE.UNIT_CFG,
				iq_aeOpMode			:= fbModeSwitch.q_aeOpMode,
				iq_abOutputReady	:= fbOutputReady.q_abReady,
				iq_astUnitP			:= fbAutoGate.q_astUnitP,
				iq_astUnitQ			:= fbAutoGate.q_astUnitQ,
				iq_astGrpP			:= fbAutoGate.q_astGrpP,
				iq_astGrpQ			:= fbAutoGate.q_astGrpQ,
				iq_astGrpPLim		:= fbSelect.q_astAutoGrpPLim,
				iq_astGrpQLim		:= fbSelect.q_astAutoGrpQLim,
				iq_afOtherGrpP		:= fbManualShape.q_afGrpP,
				iq_afOtherGrpQ		:= fbManualShape.q_afGrpQ,
				iq_aabLimOn			:= fbLimitEval.q_aabOn,
				iq_aastLim			:= fbLimitEval.q_aastLim,
				iq_aaeBasis			:= fbLimitEval.q_aaeBasis,
				iq_aanLimModule		:= fbLimitEval.q_aanModule,
				iq_abPccManual		:= fbLimitEval.q_abPccManual,
				iq_abResume			:= fbLimitEval.q_abResume,
				iq_afPComp			:= fbLimitEval.q_afPComp,
				iq_afQComp	:= fbLimitEval.q_afQComp,
				iq_astGroupEnv	:= fbEquipLimits.q_astGroupEnv);

(* ===== 5. [제어 그룹마다] 유닛 한도 · 분배 ===== *)
fbDistributor(	iq_aipDistPolicy	:= GVL_SITE.g_aipDistPolicy,
				iq_afAutoGrpP		:= fbAutoShape.q_afGrpP,
				iq_afAutoGrpQ		:= fbAutoShape.q_afGrpQ,
				iq_afAutoUnitP		:= fbAutoShape.q_afUnitP,
				iq_afAutoUnitQ		:= fbAutoShape.q_afUnitQ,
				iq_astAutoUnitP		:= fbAutoGate.q_astUnitP,
				iq_astAutoUnitQ		:= fbAutoGate.q_astUnitQ,
				iq_abAutoGrpPCmd	:= fbAutoShape.q_abGrpPCmd,
				iq_abAutoGrpQCmd	:= fbAutoShape.q_abGrpQCmd,
				iq_afManualGrpP		:= fbManualShape.q_afGrpP,
				iq_afManualGrpQ		:= fbManualShape.q_afGrpQ,
				iq_afManualUnitP	:= fbManualShape.q_afUnitP,
				iq_afManualUnitQ	:= fbManualShape.q_afUnitQ,
				iq_astManualUnitP	:= fbManualGate.q_astUnitP,
				iq_astManualUnitQ	:= fbManualGate.q_astUnitQ,
				iq_abManualGrpPCmd	:= fbManualShape.q_abGrpPCmd,
				iq_abManualGrpQCmd	:= fbManualShape.q_abGrpQCmd,
				iq_astManualPolicy	:= GVL_PERSIST.g_astManualPolicy,
				iq_aeOpMode			:= fbModeSwitch.q_aeOpMode,
				iq_astUnitEnv	:= fbEquipLimits.q_astUnitEnv,
				iq_astBatEnv	:= fbEquipLimits.q_astBatEnv,
				iq_astUnitCfg	:= GVL_SITE.UNIT_CFG,
				iq_astBatGroup	:= fbBatGroup.q_astBatGroup,
				iq_astGroupSet	:= GVL_PERSIST.g_astGroupSet,
				iq_abOutputReady	:= fbOutputReady.q_abReady,
				iq_aeNotReadyBy	:= fbOutputReady.q_aeNotReadyBy);

(* ===== 6. 쓰기 (시퀀서 · 디스패처) ===== *)
fbSequencer(	i_bTestReset	:= bTestReset,
				i_bCmdEnable	:= fbConfigCheck.q_bConfigOk,
				i_bWriteEnable	:= bWriteEnable,
				iq_abNewReq		:= fbStateArb.q_abNewReq,
				iq_aeReq		:= fbStateArb.q_aeReq,
				iq_astUnitProt	:= fbProtection.q_astUnitProt,
				iq_aeStartMode	:= GVL_SITE.START_MODE,
				iq_astUnit		:= fbSnapshot.q_astUnit,
				iq_astAvail		:= fbUnitAvail.q_astAvail,
				iq_astUnitCfg	:= GVL_SITE.UNIT_CFG,
				iq_astBms		:= fbSnapshot.q_astBms,
				iq_astBmsCfg	:= GVL_SITE.BMS_CFG,
				iq_astBmsAvail	:= fbBatGroup.q_astBmsAvail,
				iq_astBmsProt	:= fbProtection.q_astBmsProt,
				iq_astSrcOut	:= fbSources.q_astOut,
				iq_astReg		:= GVL_PERSIST.g_astSourceReg,
				iq_aeOpMode		:= fbModeSwitch.q_aeOpMode,
				iq_stSet		:= GVL_PERSIST.g_stSeqSet);

// 그룹 상태 요약 (그룹 보기에 다음 스캔부터)
fbGroupState(	iq_aeUnitSeq	:= fbSequencer.q_aeUnitSeq,
				iq_astUnitCfg	:= GVL_SITE.UNIT_CFG);

fbDispatcher(	i_tWritePeriod	:= GVL_PERSIST.g_stSeqSet.tWritePeriod,
				i_bWriteEnable	:= bWriteEnable,
				iq_aipPcs		:= GVL_SITE.g_aipPcs,
				iq_aipBms		:= GVL_SITE.g_aipBms,
				iq_astUnitCfg	:= GVL_SITE.UNIT_CFG,
				iq_astUnitCmd	:= fbSequencer.q_astUnitCmd,
				iq_abOutputReady	:= fbOutputReady.q_abReady,
				iq_astUnitSet	:= fbDistributor.q_astUnitSet,
				iq_astBmsCmd	:= fbSequencer.q_astBmsCmd,
				iq_aeOpMode		:= fbModeSwitch.q_aeOpMode,
				iq_abManualNew	:= fbManualGate.q_abNew,
				iq_abManualFollow:= fbManualShape.q_abFollow,
				iq_abUnitLimited:= fbDistributor.q_abUnitLimited);

// 보조 장비 출력(DO): 출력 규칙 → 지연·유지 → 같은 점은 OR (DO는 여기서만 씀)
fbAuxOutput(	i_bReset		:= bClearHoldDo,
				i_bWriteEnable	:= bWriteEnable,
				iq_astCfg		:= GVL_PERSIST.g_astOutputCfg,
				iq_aipRule		:= GVL_SITE.g_aipOutput,
				iq_aipAux		:= GVL_SITE.g_aipAux);

(* ===== 옆: 출력 진단 · 이벤트 로그 · 보고 ===== *)

fbAlive(		iq_nLastAlive	:= GVL_PERSIST.g_nLastAliveLocal,
				iq_sLastAlive	:= GVL_PERSIST.g_sLastAlive);

// PERSISTENT 저장: 운영 설정이 바뀌면 1 s 뒤 바로, 그리고 주기마다 (GVL_PERSIST에 설정을 추가하면 여기도 연결)
fbPersistSave(	i_tPeriod		:= GVL_SITE.LOG_SET.tPersistSave,
				i_bSaveNow		:= fbUpsConfigApply[1].q_bDesiredChanged OR fbUpsCommand[1].q_bDesiredChanged OR fbBmsRack[1].q_bMaskChanged,	// UPS 설정 보관값이 바뀌면 바로 저장 (CF-UPS-02)
				iq_aeOpMode		:= GVL_PERSIST.g_aeOpMode,
				iq_astGroupSet	:= GVL_PERSIST.g_astGroupSet,
				iq_astManualPolicy:= GVL_PERSIST.g_astManualPolicy,
				iq_astSourceReg	:= GVL_PERSIST.g_astSourceReg,
				iq_astLimitReg	:= GVL_PERSIST.g_astLimitReg,
				iq_astPermitReg	:= GVL_PERSIST.g_astPermitReg,
				iq_astCompReg	:= GVL_PERSIST.g_astCompReg,
				iq_astRuleCfg	:= GVL_PERSIST.g_astRuleCfg,
				iq_astOutputCfg	:= GVL_PERSIST.g_astOutputCfg,
				iq_astUnitRuleReg	:= GVL_PERSIST.g_astUnitRuleReg,
				iq_astBatRuleReg	:= GVL_PERSIST.g_astBatRuleReg,
				iq_stCmdFilter	:= GVL_PERSIST.g_stCmdFilter,
				iq_stManualCmdSet	:= GVL_PERSIST.g_stManualCmdSet,
				iq_stSeqSet		:= GVL_PERSIST.g_stSeqSet,
				iq_stBrokerWatch	:= GVL_PERSIST.g_stBrokerWatch,	// [9번 수정 2026-11-09: 추가]
				i_pModuleSet	:= ADR(GVL_PERSIST.g_stModuleSet),
				i_nModuleSetSize	:= SIZEOF(GVL_PERSIST.g_stModuleSet));

fbOutputDiag(	iq_astAutoShape		:= fbAutoShape.q_astDiag,
				iq_astManualShape	:= fbManualShape.q_astDiag,
				iq_astDist		:= fbDistributor.q_astDistDiag,
				iq_astUnitDiag	:= fbDistributor.q_astUnitDiag,
				iq_aeOpMode		:= fbModeSwitch.q_aeOpMode,
				iq_aeGroupState	:= fbGroupState.q_aeGroupState,
				iq_astWritten	:= fbDispatcher.q_astWritten,
				iq_astUnitSet	:= fbDistributor.q_astUnitSet,
				iq_astUnitCfg	:= GVL_SITE.UNIT_CFG);

fbEventLog(		i_stSet			:= GVL_SITE.LOG_SET,
				i_bTestMode		:= GVL_SITE.TEST_MODE,
				i_nConfigErrors	:= fbConfigCheck.q_nErrors,
				iq_asConfigErrors	:= fbConfigCheck.q_asErrors,
				i_bSetChanged	:= fbPersistSave.q_bSetChanged OR fbEmsCfg.q_bApplied,	// [9-21 수정 2026-11-04: EMS config 반영도 기록. 원래 fbPersistSave.q_bSetChanged]
				i_sSetChanged	:= SEL(fbEmsCfg.q_bApplied, fbPersistSave.q_sSetChanged, fbEmsCfg.q_sApplied),	// [9-21 수정 2026-11-04: 원래 fbPersistSave.q_sSetChanged]
				i_bSetRejected	:= fbSettingGuard.q_bRejected OR fbEmsCfg.q_bRejected,	// [9-21 수정 2026-11-04: EMS config 거부도 기록. 원래 fbSettingGuard.q_bRejected]
				i_sSetRejected	:= SEL(fbSettingGuard.q_bRejected, fbEmsCfg.q_sRejected, fbSettingGuard.q_sRejected),	// [9-21 수정 2026-11-04: 원래 fbSettingGuard.q_sRejected]
				i_bPersistError	:= fbPersistSave.q_bError,
				i_nPersistErrorId	:= fbPersistSave.q_nErrorId,
				i_bPmsStart		:= fbAlive.q_bStartEvent,
				i_sStartLastAlive	:= fbAlive.q_sLastAlive,
				i_sStartOffTime	:= fbAlive.q_sOffTime,
				i_bRedUse		:= GVL_SITE.RED_SET.bUse,
				i_eRedRole		:= GVL_IF.g_eRedRole,
				i_eRedState		:= GVL_IF.g_eRedState,
				i_ePeer			:= GVL_IF.g_ePeerState,
				i_nSwitchCount	:= GVL_IF.g_nRedSwitchCount,
				i_eSwitch		:= GVL_IF.g_eRedSwitch,
				i_nResumeCount	:= GVL_IF.g_nRedResumeCount,
				i_nSyncApplied	:= GVL_IF.g_nSyncApplied,
				i_bSyncFresh	:= GVL_IF.g_bSyncFresh,
				i_bPeerEapOk	:= GVL_IF.g_bPeerEapOk,
				i_bRoleConflict	:= GVL_IF.g_bRedRoleConflict,
				i_bBrokerLost	:= fbBrokerWatch.q_bLost,		// [9번 수정 2026-11-09: 추가]
				i_sBrokerName	:= fbBrokerWatch.q_sBroker,
				i_sBrokerDelay	:= fbBrokerWatch.q_sDelay,
				iq_aabRule		:= fbProtection.q_aabRule,
				iq_astRuleCfg	:= GVL_PERSIST.g_astRuleCfg,
				iq_aeUnitSeq	:= fbSequencer.q_aeUnitSeq,
				iq_aeRefuse		:= fbSequencer.q_aeRefuse,
				iq_aeBatRefuse	:= fbSequencer.q_aeBatRefuse,
				iq_abBatRefusedNow:= fbSequencer.q_abBatRefusedNow,
				iq_aeFailCmd	:= fbSequencer.q_aeFailCmd,
				iq_aeBmsFailCmd	:= fbSequencer.q_aeBmsFailCmd,
				iq_aeOpMode		:= fbModeSwitch.q_aeOpMode,
				iq_abModeForced	:= fbModeSwitch.q_abModeForced,
				iq_astUnitProt	:= fbProtection.q_astUnitProt,
				iq_abBadValue	:= fbSelect.q_abBadValue,
				iq_afBadValue	:= fbSelect.q_afBadValue,
				iq_aeManualRefuse	:= fbManualGate.q_aeRefuse,
				iq_anManualRefuseModule:= fbManualGate.q_anRefuseModule,
				iq_astSrcOut	:= fbSources.q_astOut,
				iq_abPcsReqTaken:= fbStateArb.q_abPcsReqTaken,
				iq_abBatReqTaken:= fbSequencer.q_abBatReqTaken,
				iq_astReg		:= GVL_PERSIST.g_astSourceReg,
				iq_astAutoPDiag	:= fbOutputDiag.q_astAutoPDiag,
				iq_astUnitDiag	:= fbDistributor.q_astUnitDiag,
				iq_astVirtual	:= GVL_TEST.g_astVirtual,
				iq_abBadSet		:= fbDispatcher.q_abBadSet,
				iq_abWaitPermit	:= fbSequencer.q_abWaitPermit,
				iq_abPermit		:= fbPermitEval.q_abPermit,
				iq_anPermitModule	:= fbPermitEval.q_anPermitModule,
				iq_anPermitReason	:= fbPermitEval.q_anPermitReason,
				iq_astUnit		:= fbSnapshot.q_astUnit,
				iq_astBms		:= fbSnapshot.q_astBms,
				iq_aipRule		:= GVL_SITE.g_aipRule,
				iq_aipResp		:= GVL_SITE.g_aipResp,	// [결함 8 수정 2026-11-03: 추가]
				iq_aipSource	:= GVL_SITE.g_aipSource,
				iq_aipModule	:= fbModuleList.q_aipModule,
				iq_fbCtrlMode	:= GVL_SITE.g_fbCtrlMode1);	// [7번 수정 2026-11-09: 제어 모드 전환·거부·스스로 끝남 기록]

fbReport(		iq_astUnit		:= fbSnapshot.q_astUnit,
				iq_astBms		:= fbSnapshot.q_astBms,
				iq_astView		:= fbGroupView.q_astView,
				iq_astAutoPDiag	:= fbOutputDiag.q_astAutoPDiag,
				iq_aeUnitSeq	:= fbSequencer.q_aeUnitSeq,
				iq_astWritten	:= fbDispatcher.q_astWritten);

// BMS 랙 컨택터 개별 제어 (EMS command/bat 11·12). 일괄(1·2)은 코어 경로. 쓰기 막힘·허가·통신은 드라이버가 판단
fbBmsRack[1](i_stCmd:=GVL_SITE.g_fbSrcEms.i_stCmd.astBatRack[1], i_nRackCount:=GVL_PARAM.RACKS_PER_BMS,
 i_wRestore:=GVL_PERSIST.g_awBmsRackMask[1], i_bAccepted:=abBmsRackAcc[1], i_eDriverResult:=aeBmsRackRes[1],
 i_wActual:=GVL_SITE.g_fbBms1.q_stState.wRackContactor, i_bActualValid:=GVL_SITE.g_fbBms1.q_stState.bContactorFeedbackKnown);
abBmsRackAcc[1]:=FALSE; aeBmsRackRes[1]:=E_UpsResult.None;
IF fbBmsRack[1].q_bWriteReq THEN
 abBmsRackAcc[1]:=GVL_SITE.g_fbBms1.M_SetRackMask(i_wMask:=fbBmsRack[1].q_wWriteMask);
 aeBmsRackRes[1]:=GVL_SITE.g_fbBms1.q_eRequestResult;
END_IF
GVL_PERSIST.g_awBmsRackMask[1]:=fbBmsRack[1].q_wMask;

// BMS 컨택터 하나씩 제어 (EMS command/bat 5~10: 40013 랙 전체, 40014 충전, 40015 방전) [2026-11-13]
// 11·12처럼 코어 순서(유닛 정지 확인)를 거치지 않음. 쓰기 막힘·허가·통신은 드라이버가 판단
fbBmsCtl[1](i_stCmd:=GVL_SITE.g_fbSrcEms.i_stCmd.astBatCtl[1], i_bAccepted:=abBmsCtlAcc[1], i_eDriverResult:=aeBmsCtlRes[1]);
abBmsCtlAcc[1]:=FALSE; aeBmsCtlRes[1]:=E_UpsResult.None;
IF fbBmsCtl[1].q_bWriteReq THEN
 abBmsCtlAcc[1]:=GVL_SITE.g_fbBms1.M_SetControl(i_eControl:=fbBmsCtl[1].q_eControl, i_bOn:=fbBmsCtl[1].q_bOn);
 aeBmsCtlRes[1]:=GVL_SITE.g_fbBms1.q_eRequestResult;
END_IF

// BMS 쓰기 시험: 코어 경로와 별개인 시험 명령. 접수 뒤 전송은 드라이버 M_Cycle이 함
IF nBmsTestCmd <> 0 THEN
 CASE nBmsTestCmd OF
  1: GVL_SITE.g_fbBms1.M_SetRackMask(i_wMask := wBmsTestValue);
  2: GVL_SITE.g_fbBms1.M_SetControl(i_eControl := E_EsolutionControl.ChargeContactor, i_bOn := bBmsTestOn);
  3: GVL_SITE.g_fbBms1.M_SetControl(i_eControl := E_EsolutionControl.DischargeContactor, i_bOn := bBmsTestOn);
  4: GVL_SITE.g_fbBms1.M_SetControl(i_eControl := E_EsolutionControl.SystemContactor, i_bOn := bBmsTestOn);
  5: GVL_SITE.g_fbBms1.M_SetControl(i_eControl := E_EsolutionControl.EmergencyShutdown, i_bOn := TRUE);
  6:
   nBmsTestSeq := nBmsTestSeq + 1;
   stBmsTestCmd.eCmd := E_BatCmd.Reset;
   stBmsTestCmd.nSeq := nBmsTestSeq;
   GVL_SITE.g_fbBms1.M_SetStateCmd(i_stCmd := stBmsTestCmd);
  7: GVL_SITE.g_fbBms1.M_RequestOperation(i_eOperation := E_EsolutionOperation.PeriodicStart);
  8: GVL_SITE.g_fbBms1.M_RequestOperation(i_eOperation := E_EsolutionOperation.DischargeCancel);
 END_CASE
 eBmsTestResult := GVL_SITE.g_fbBms1.q_eRequestResult;
 nBmsTestCmd := 0;
END_IF

// 충방전 요청 생성. 실제 장비 쓰기에는 연결하지 않음.
// 통신 시험 중 충방전 알고리즘 호출 중지 (2026-11-02)
//afbUpsCharge[1](i_bEnable:=GVL_PARAM.UPS_ALGORITHM_ENABLED AND abUpsChargeEnable[1],
// i_bCancel:=abUpsChargeCancel[1], i_bReset:=abUpsChargeReset[1], i_eMode:=aeUpsChargeMode[1],
// i_stSet:=astUpsChargeSet[1], i_stUps:=GVL_SITE.g_fbUps1.q_stState,
// i_stBms:=GVL_SITE.g_fbBms1.q_stState, i_stTime:=fbClock.q_stTime, i_stFeedback:=astUpsChargeFeedback[1]);
//afbUpsTemp[1](i_bEnable:=GVL_PARAM.UPS_ALGORITHM_ENABLED AND abUpsTempEnable[1],
// i_bSuspend:=(afbUpsCharge[1].q_eMode = E_UpsChargeMode.Periodic OR afbUpsCharge[1].q_eMode = E_UpsChargeMode.Pulse)
// AND afbUpsCharge[1].q_eStep >= E_UpsChargeStep.PrepareBms AND afbUpsCharge[1].q_eStep <= E_UpsChargeStep.CancelBms,
// i_bReset:=abUpsChargeReset[1], i_stUps:=GVL_SITE.g_fbUps1.q_stState,
// i_stSet:=astUpsChargeSet[1], i_stTime:=fbClock.q_stTime, i_stFeedback:=astUpsTempFeedback[1]);
A_Report();

ACTION A_PassModuleSet:
// 모듈 설정 넘기기: GVL_PERSIST.g_stModuleSet 칸 → 모듈 i_stSet. 현장 모듈마다 한 줄 (운전 중 바꾼 값이 이 스캔부터 적용)
GVL_SITE.g_fbSocLimit.i_stSet	:= GVL_PERSIST.g_stModuleSet.stSocLimit;
// 제어 모드: 접속점 그룹 관리자에 모드 등록 배열·설정·시각·유닛 값 주소(유닛 단위일 때만 씀), 모드마다 설정 (공통 stCmCommon은 같이 씀)
GVL_SITE.g_fbCtrlMode1.i_aipMode	:= GVL_SITE.g_aipCtrlMode1;
GVL_SITE.g_fbCtrlMode1.i_stSet	:= GVL_PERSIST.g_stModuleSet.stCtrlMode1;
GVL_SITE.g_fbCtrlMode1.i_stTime	:= fbClock.q_stTime;
GVL_SITE.g_fbCtrlMode1.i_pUnitView	:= ADR(fbUnitView.q_astView);
GVL_SITE.g_fbCmConstP1.i_stSet	:= GVL_PERSIST.g_stModuleSet.stCmConstP1;
GVL_SITE.g_fbCmSchedule1.i_stCommon	:= GVL_PERSIST.g_stModuleSet.stCmCommon;
GVL_SITE.g_fbCmSchedule1.i_stTable	:= GVL_PERSIST.g_stModuleSet.stCmSchedule1;
GVL_SITE.g_fbCmPeakCut1.i_stCommon	:= GVL_PERSIST.g_stModuleSet.stCmCommon;
GVL_SITE.g_fbCmPeakCut1.i_stSet	:= GVL_PERSIST.g_stModuleSet.stCmPeakCut1;
GVL_SITE.g_fbCmSchedPeak1.i_stCommon	:= GVL_PERSIST.g_stModuleSet.stCmCommon;
GVL_SITE.g_fbCmSchedPeak1.i_stTable	:= GVL_PERSIST.g_stModuleSet.stCmSchedule1;
GVL_SITE.g_fbCmSchedPeak1.i_stSet	:= GVL_PERSIST.g_stModuleSet.stCmSchedPeak1;
// [16번 수정 2026-11-09: 관리자 PCS2(g_fbCtrlMode2)와 모드 두 번째 세트 줄 없앰]
GVL_SITE.g_fbUnitLimit.i_stSet	:= GVL_PERSIST.g_stModuleSet.stUnitLimit;	// [9-21 수정 2026-11-04: 사용자 한도 기본 등록. 원래 주석 예 "// 예: GVL_SITE.g_fbUnitLimit.i_stSet := GVL_PERSIST.g_stModuleSet.stUnitLimit;"]
END_ACTION

ACTION A_PassEmsCfg:
// [9-21 수정 2026-11-04: 추가] EMS config 받기: GVL_IF.g_stEmsCfg를 번호를 확인하며 복사해 FB_EmsConfigApply에 넘김 (A_PassEmsCmd와 같은 읽는 규칙)
// 쓰는 곳은 GVL_PERSIST 모듈 설정(영속). 실제 설정 echo는 본문에서 설정 보호 뒤에 GVL_IF.g_stEmsCfgEcho에 씀
nEmsCfgSeq := GVL_IF.g_nCfgSeq;
bEmsCfgOk := FALSE;
IF (nEmsCfgSeq AND 1) = 0 THEN
	stEmsCfgCopy := GVL_IF.g_stEmsCfg;
	bEmsCfgOk := GVL_IF.g_nCfgSeq = nEmsCfgSeq;
END_IF
fbEmsCfg(	i_bValid		:= bEmsCfgOk,
			i_stCfg			:= stEmsCfgCopy,
			i_astUnitCfg	:= GVL_SITE.UNIT_CFG,
			iq_stSocLimit	:= GVL_PERSIST.g_stModuleSet.stSocLimit,
			iq_stUnitLimit	:= GVL_PERSIST.g_stModuleSet.stUnitLimit);
END_ACTION

